q_bDone := FALSE;
q_bError := FALSE;
_bStartInput := FALSE; _bStartHolding := FALSE; _bStartWrite := FALSE; _bStartMulti := FALSE;
_rtExecute(CLK := i_bExecute);
IF _rtExecute.Q AND NOT q_bBusy THEN
	q_nErrorId := 0;
	IF i_sIpAddr = '' OR i_nPort = 0 OR i_nQuantity = 0 OR i_nQuantity > 125 THEN
		q_bDone := TRUE; q_bError := TRUE; q_nErrorId := 16#F001;
	ELSIF (i_nFunction = 6 AND (NOT GVL_PARAM.UPS_CONTROL_ENABLED OR NOT i_bWritePermit OR i_nQuantity <> 1))
		OR (i_nFunction = 16 AND (NOT GVL_PARAM.UPS_CONTROL_ENABLED OR NOT i_bWritePermit OR i_nQuantity > 3)) THEN
		q_bDone := TRUE; q_bError := TRUE; q_nErrorId := 16#F002;
	ELSIF i_nFunction <> 3 AND i_nFunction <> 4 AND i_nFunction <> 6 AND i_nFunction <> 16 THEN
		q_bDone := TRUE; q_bError := TRUE; q_nErrorId := 16#F003;
	ELSE
		_sIpAddr:=i_sIpAddr; _nPort:=i_nPort; _nUnitId:=i_nUnitId;
		_tTimeout:=i_tTimeout; _nAddress:=i_nAddress; _wValue:=i_wValue; _awValues:=i_awValues;
		_nFunction := i_nFunction; _nQuantity := i_nQuantity; q_bBusy := TRUE;
		_bStartInput := _nFunction = 4; _bStartHolding := _nFunction = 3; _bStartWrite := _nFunction = 6;
		_bStartMulti := _nFunction = 16;
	END_IF
END_IF
// Call all instances every scan, also while disabled, to drain an in-flight transaction.
_fbInput(sIPAddr:=_sIpAddr,nTCPPort:=_nPort,nUnitID:=_nUnitId,nMBAddr:=_nAddress,nQuantity:=_nQuantity,
	cbLength:=SIZEOF(q_awData),pDestAddr:=ADR(q_awData),tTimeout:=_tTimeout,bExecute:=_bStartInput);
_fbHolding(sIPAddr:=_sIpAddr,nTCPPort:=_nPort,nUnitID:=_nUnitId,nMBAddr:=_nAddress,nQuantity:=_nQuantity,
	cbLength:=SIZEOF(q_awData),pDestAddr:=ADR(q_awData),tTimeout:=_tTimeout,bExecute:=_bStartHolding);
_fbSingle(sIPAddr:=_sIpAddr,nTCPPort:=_nPort,nUnitID:=_nUnitId,nMBAddr:=_nAddress,nValue:=_wValue,tTimeout:=_tTimeout,bExecute:=_bStartWrite);
_fbMulti(sIPAddr:=_sIpAddr,nTCPPort:=_nPort,nUnitID:=_nUnitId,nQuantity:=_nQuantity,nMBAddr:=_nAddress,
	cbLength:=WORD_TO_UDINT(_nQuantity)*2,pSrcAddr:=ADR(_awValues),tTimeout:=_tTimeout,bExecute:=_bStartMulti);
IF q_bBusy THEN
	CASE _nFunction OF
		4: IF NOT _fbInput.bBusy AND NOT _bStartInput THEN
				q_bDone := TRUE; q_bError := _fbInput.bError OR (_fbInput.cbRead <> WORD_TO_UDINT(_nQuantity)*2);
				q_nErrorId := _fbInput.nErrId; q_bBusy := FALSE; END_IF
		3: IF NOT _fbHolding.bBusy AND NOT _bStartHolding THEN
				q_bDone := TRUE; q_bError := _fbHolding.bError OR (_fbHolding.cbRead <> WORD_TO_UDINT(_nQuantity)*2);
				q_nErrorId := _fbHolding.nErrId; q_bBusy := FALSE; END_IF
		6: IF NOT _fbSingle.bBusy AND NOT _bStartWrite THEN
				q_bDone := TRUE; q_bError := _fbSingle.bError; q_nErrorId := _fbSingle.nErrId; q_bBusy := FALSE; END_IF
		16: IF NOT _fbMulti.bBusy AND NOT _bStartMulti THEN
				q_bDone := TRUE; q_bError := _fbMulti.bError; q_nErrorId := _fbMulti.nErrId; q_bBusy := FALSE; END_IF
	END_CASE
	IF q_bDone AND q_bError AND q_nErrorId = 0 THEN q_nErrorId := 16#F004; END_IF
END_IF

END_FUNCTION_BLOCK

// ---- 20_Module/Ups/F_UpsNextSeq.TcPOU
FUNCTION F_UpsNextSeq : UDINT
VAR_INPUT i_nSeq : UDINT; END_VAR

IF i_nSeq = 16#FFFFFFFF THEN F_UpsNextSeq := 1;
ELSE F_UpsNextSeq := i_nSeq + 1; END_IF

END_FUNCTION

// ---- 20_Module/Virtual/FB_MeterSim.TcPOU
FUNCTION_BLOCK FB_MeterSim EXTENDS FB_DeviceBase IMPLEMENTS I_Meter		// 가상 계측기 (시험용)
VAR_INPUT
	i_fP			: REAL;					// kW (방전 +). PRG_SimLink가 넣음
	i_fQ			: REAL;					// kvar
	i_fVPhase		: REAL := 13221.0;		// V, 상전압
	i_fHz			: REAL := 60.0;
	i_bForceInvalid	: BOOL;			// 시험: 접속점 P/Q 계측 무효 (값·통신·전압·주파수는 유지)
END_VAR
VAR
	_stMeter		: ST_MeterState;
END_VAR

PROPERTY MeterState : ST_MeterState
GET
MeterState := _stMeter;
END_GET
END_PROPERTY

METHOD M_Cycle
VAR
	k		: UINT;
END_VAR
IF M_IsReadTime() THEN		// 읽기 주기마다 응답한 것으로 봄
	M_MarkAlive();
END_IF
M_UpdateComm();

_stMeter.bComm			:= _bComm;
_stMeter.stP.fValue		:= i_fP;
_stMeter.stP.bValid		:= NOT i_bForceInvalid;
_stMeter.stQ.fValue		:= i_fQ;
_stMeter.stQ.bValid		:= NOT i_bForceInvalid;
_stMeter.stV.fValue		:= i_fVPhase;
_stMeter.stV.bValid		:= TRUE;
FOR k := 1 TO 3 DO
	_stMeter.astV[k].fValue	:= i_fVPhase;
	_stMeter.astV[k].bValid	:= TRUE;
END_FOR
_stMeter.stF.fValue		:= i_fHz;
_stMeter.stF.bValid		:= TRUE;
END_METHOD

END_FUNCTION_BLOCK

// ---- 20_Module/Driver/Sebang/FB_SebangUps.TcPOU
FUNCTION_BLOCK FB_SebangUps EXTENDS FB_DeviceBase IMPLEMENTS I_Ups

VAR_INPUT
	i_bEnable : BOOL;
	i_sIpAddr : STRING(15);
	i_nPort : UINT := 502;
	i_nUnitId : BYTE := 1;
	i_tTimeout : TIME := T#1S;
	i_bWritePermit : BOOL; // site dispatcher: config OK AND active PLC
	i_bBlockStart : BOOL; // 2026-11-17: UPS 고장·e-stop 중 (MAIN이 보고 Status b2 OR b3로 줌). 시작 명령·설정 쓰기를 대기열에 넣지 않고, 이미 들어간 것도 뺌
END_VAR
VAR_OUTPUT
	q_eRequestResult : E_UpsResult;
	q_nTransportError : UDINT;
END_VAR
VAR
	_fbJob : FB_UpsModbusJob;
	_bLaunch : BOOL;
	_bCurrentWrite : BOOL;
	_bDiscardResponse : BOOL; // response started before a disable must not complete a new snapshot
	_nFunction : UINT;
	_nAddress : WORD;
	_nQuantity : WORD;
	_wValue : WORD;
	_bPendingWrite : BOOL;
	_nPendingAddress : WORD;
	_wPendingValue : WORD;
	_nPoll : UINT;
	_nCopy : UINT;
	_bReadDue : BOOL;
	_bCycle : BOOL; // 2026-11-23 한 바퀴(요청 4개) 읽는 중. i_tReadPeriod마다 시작해 4개를 연달아 읽음 (명세 DV-04 v2.46)
END_VAR

VAR_OUTPUT
	q_stRaw : ST_UpsRaw;
	q_stState : ST_UpsState;
END_VAR
VAR
	_stWork : ST_UpsRaw;
	_nSampleSeq : UDINT;
END_VAR

METHOD M_Cycle
_bReadDue := M_IsReadTime();
IF _bReadDue THEN _bCycle:=TRUE; END_IF // 한 바퀴 시작 (명세 DV-04 v2.46: 주기 = 한 바퀴)
IF NOT i_bEnable THEN
	_bDiscardResponse:=_bDiscardResponse OR _fbJob.q_bBusy;
	_bLaunch:=FALSE;
END_IF
IF NOT i_bEnable OR NOT i_bWritePermit OR NOT GVL_PARAM.UPS_CONTROL_ENABLED THEN
	_bPendingWrite := FALSE;
	// A queued but not yet started FC06 must not survive a gate transition.
	IF _bLaunch AND _bCurrentWrite THEN _bLaunch := FALSE; END_IF
END_IF
// 2026-11-17: 대기 중에 고장·e-stop이 생기면 시작 명령(켜기·시작)과 설정 쓰기를 뺀다. 끄기·취소·리셋(101,103,105,107,109,113,117,119,121,123,125,100)은 그대로
IF i_bBlockStart THEN
	IF _bPendingWrite THEN
		CASE _nPendingAddress OF
			7..64, 102, 104, 106, 108, 110, 111, 112, 114, 115, 116, 118, 120, 122, 124:
				_bPendingWrite := FALSE;
				q_eRequestResult := E_UpsResult.BadRequest;
		END_CASE
	END_IF
	IF _bLaunch AND _bCurrentWrite THEN
		CASE _nAddress OF
			7..64, 102, 104, 106, 108, 110, 111, 112, 114, 115, 116, 118, 120, 122, 124:
				_bLaunch := FALSE;
				_bCurrentWrite := FALSE;
				q_eRequestResult := E_UpsResult.BadRequest;
		END_CASE
	END_IF
END_IF
_fbJob(i_sIpAddr:=i_sIpAddr,i_nPort:=i_nPort,i_nUnitId:=i_nUnitId,i_tTimeout:=i_tTimeout,
	i_bExecute:=_bLaunch,i_bWritePermit:=i_bWritePermit AND i_bEnable,
	i_nFunction:=_nFunction,i_nAddress:=_nAddress,i_nQuantity:=_nQuantity,i_wValue:=_wValue);
_bLaunch := FALSE;
IF _fbJob.q_bDone THEN
	q_nTransportError := _fbJob.q_nErrorId;
	IF _bCurrentWrite THEN M_MarkWriteResult(NOT _fbJob.q_bError); END_IF
END_IF

IF _fbJob.q_bDone AND _bDiscardResponse THEN
	_bDiscardResponse:=FALSE; _nPoll:=0; _bCycle:=FALSE;
ELSIF _fbJob.q_bDone AND NOT _bCurrentWrite THEN
	IF _fbJob.q_bError THEN _nPoll:=0; _bCycle:=FALSE; // 다음 주기에 처음부터
	ELSE
		CASE _nPoll OF
			0: FOR _nCopy:=0 TO 34 DO _stWork.awInput[_nCopy]:=_fbJob.q_awData[_nCopy]; END_FOR
			1: FOR _nCopy:=0 TO 15 DO _stWork.awInput[_nCopy+38]:=_fbJob.q_awData[_nCopy]; END_FOR
			2: FOR _nCopy:=0 TO 11 DO _stWork.awParam[_nCopy]:=_fbJob.q_awData[_nCopy]; END_FOR
			3: FOR _nCopy:=0 TO 16 DO _stWork.awParam[_nCopy+50]:=_fbJob.q_awData[_nCopy]; END_FOR
		END_CASE
		IF _nPoll=3 THEN
			q_stRaw:=_stWork; _nSampleSeq:=F_UpsNextSeq(_nSampleSeq); M_MarkAlive(); _nPoll:=0; _bCycle:=FALSE;
		ELSE _nPoll:=_nPoll+1; END_IF
	END_IF
END_IF
M_UpdateComm();
q_stState:=F_DecodeSebangUps(q_stRaw);
q_stState.bComm:=_bComm AND i_bEnable;
q_stState.bValid:=q_stState.bComm AND _nSampleSeq<>0;
q_stState.nSampleSeq:=_nSampleSeq;
q_stState.bWriteFail:=_bWriteFail;
IF NOT _fbJob.q_bBusy AND NOT _fbJob.q_bDone AND i_bEnable AND i_sIpAddr<>'' THEN
IF _bPendingWrite THEN
	_nFunction:=6; _nAddress:=_nPendingAddress; _nQuantity:=1; _wValue:=_wPendingValue;
	_bCurrentWrite:=TRUE; _bPendingWrite:=FALSE; _bLaunch:=TRUE;
ELSIF _bCycle THEN // 한 바퀴 안에서는 앞 요청이 끝나면 바로 다음 요청 (쓰기가 있으면 쓰기 먼저)
	_bCurrentWrite:=FALSE;

	CASE _nPoll OF
		0: _nFunction:=4; _nAddress:=0; _nQuantity:=35;
		1: _nFunction:=4; _nAddress:=38; _nQuantity:=16;
		2: _nFunction:=3; _nAddress:=0; _nQuantity:=12;
		3: _nFunction:=3; _nAddress:=50; _nQuantity:=17;
	END_CASE
	_bLaunch:=TRUE;
	END_IF
END_IF
IF NOT i_bEnable THEN _nSampleSeq:=0; _nPoll:=0; _bLaunch:=FALSE; _bCycle:=FALSE; END_IF
END_METHOD

PROPERTY UpsState : ST_UpsState
GET
UpsState:=q_stState;
END_GET
END_PROPERTY

METHOD PRIVATE M_QueueWrite : BOOL
VAR_INPUT i_nAddress : WORD; i_wValue : WORD; END_VAR
q_eRequestResult := E_UpsResult.Disabled;
IF NOT GVL_PARAM.UPS_CONTROL_ENABLED OR NOT i_bWritePermit OR NOT i_bEnable THEN RETURN; END_IF
IF i_bBlockStart THEN // 2026-11-17: 고장·e-stop 중 시작 명령·설정 쓰기는 받지 않음
	CASE i_nAddress OF
		7..64, 102, 104, 106, 108, 110, 111, 112, 114, 115, 116, 118, 120, 122, 124:
			q_eRequestResult := E_UpsResult.BadRequest;
			RETURN;
	END_CASE
END_IF
q_eRequestResult := E_UpsResult.CommUnavailable;
IF NOT _bComm THEN RETURN; END_IF
q_eRequestResult := E_UpsResult.Busy;
IF _bPendingWrite OR _bCurrentWrite AND (_fbJob.q_bBusy OR _bLaunch) THEN RETURN; END_IF
_nPendingAddress := i_nAddress; _wPendingValue := i_wValue; _bPendingWrite := TRUE;
q_eRequestResult := E_UpsResult.Accepted;
M_QueueWrite := TRUE;
END_METHOD

METHOD M_RequestCommand : BOOL
VAR_INPUT i_eCommand : E_UpsCommand; END_VAR
CASE i_eCommand OF
	E_UpsCommand.Reset,
	E_UpsCommand.BuzzerStop,
	E_UpsCommand.RectifierOn,
	E_UpsCommand.RectifierOff,
	E_UpsCommand.InverterOn,
	E_UpsCommand.InverterOff,
	E_UpsCommand.BbcOn,
	E_UpsCommand.BbcOff,
	E_UpsCommand.ToInverter,
	E_UpsCommand.ToBypass,
	E_UpsCommand.FloatCharge,
	E_UpsCommand.EqualCharge,
	E_UpsCommand.AutoOn,
	E_UpsCommand.AutoOff,
	E_UpsCommand.EmergencyDischarge,
	E_UpsCommand.PeriodicDischarge,
	E_UpsCommand.PulseDischarge,
	E_UpsCommand.CancelDischarge,
	E_UpsCommand.TrickleOn,
	E_UpsCommand.TrickleOff,
	E_UpsCommand.TemperatureOn,
	E_UpsCommand.TemperatureOff,
	E_UpsCommand.EcoOn,
	E_UpsCommand.EcoOff,
	E_UpsCommand.PrltOn,
	E_UpsCommand.PrltOff:
	M_RequestCommand:=M_QueueWrite(INT_TO_WORD(TO_INT(i_eCommand)),16#0055);
ELSE q_eRequestResult:=E_UpsResult.Unsupported;
END_CASE
END_METHOD

METHOD M_SetParameter : BOOL
// Explicit RAW register value only. 57~59 allowed since 2026-11-16 (spec v2.14: H58/H59 = voltage or SOC by H57). 62 still rejected (scale O-11).
VAR_INPUT i_nAddress : WORD; i_wRawValue : WORD; END_VAR
CASE i_nAddress OF
	7,8,10,50,51,52,53,54,55,56,57,58,59,60,61,63,64:
		M_SetParameter:=M_QueueWrite(i_nAddress,i_wRawValue);
ELSE q_eRequestResult:=E_UpsResult.Unsupported;
END_CASE
END_METHOD

METHOD M_CheckSet : WSTRING(63)
M_CheckSet:="";
IF i_bEnable THEN
	IF i_sIpAddr='' OR i_nPort=0 THEN M_CheckSet:="TCP endpoint missing";
	ELSIF i_tReadPeriod<=T#0MS OR i_tTimeout<=T#0MS OR i_tCommTimeout<=i_tReadPeriod THEN M_CheckSet:="Invalid timing";
	END_IF
END_IF
END_METHOD

END_FUNCTION_BLOCK

// ---- 20_Module/Driver/Sebang/F_DecodeSebangUps.TcPOU
FUNCTION F_DecodeSebangUps : ST_UpsState
VAR_INPUT i_stRaw : ST_UpsRaw; END_VAR
VAR n : UINT; END_VAR

// UPS Metering Data 주소 순서
F_DecodeSebangUps.fInputVoltageRV := WORD_TO_REAL(i_stRaw.awInput[0])*0.1; // 0. 입력 선간 전압 R (V)
F_DecodeSebangUps.fInputVoltageSV := WORD_TO_REAL(i_stRaw.awInput[1])*0.1; // 1. 입력 선간 전압 S (V)
F_DecodeSebangUps.fInputVoltageTV := WORD_TO_REAL(i_stRaw.awInput[2])*0.1; // 2. 입력 선간 전압 T (V)
F_DecodeSebangUps.fInputFrequencyHz := WORD_TO_REAL(i_stRaw.awInput[3])*0.1; // 3. 입력 주파수 (Hz)
F_DecodeSebangUps.fInputCurrentRA := WORD_TO_REAL(i_stRaw.awInput[4])*0.1; // 4. 입력 전류 R (A)
F_DecodeSebangUps.fInputCurrentSA := WORD_TO_REAL(i_stRaw.awInput[5])*0.1; // 5. 입력 전류 S (A)
F_DecodeSebangUps.fInputCurrentTA := WORD_TO_REAL(i_stRaw.awInput[6])*0.1; // 6. 입력 전류 T (A)
F_DecodeSebangUps.fInverterVoltageRV := WORD_TO_REAL(i_stRaw.awInput[7])*0.1; // 7. 인버터 선간 전압 R (V)
F_DecodeSebangUps.fInverterVoltageSV := WORD_TO_REAL(i_stRaw.awInput[8])*0.1; // 8. 인버터 선간 전압 S (V)
F_DecodeSebangUps.fInverterVoltageTV := WORD_TO_REAL(i_stRaw.awInput[9])*0.1; // 9. 인버터 선간 전압 T (V)
F_DecodeSebangUps.fInverterCurrentRA := WORD_TO_REAL(i_stRaw.awInput[10])*0.1; // 10. 인버터 전류 R (A)
F_DecodeSebangUps.fInverterCurrentSA := WORD_TO_REAL(i_stRaw.awInput[11])*0.1; // 11. 인버터 전류 S (A)
F_DecodeSebangUps.fInverterCurrentTA := WORD_TO_REAL(i_stRaw.awInput[12])*0.1; // 12. 인버터 전류 T (A)
F_DecodeSebangUps.fBypassVoltageRV := WORD_TO_REAL(i_stRaw.awInput[13])*0.1; // 13. 바이패스 선간 전압 R (V)
F_DecodeSebangUps.fBypassVoltageSV := WORD_TO_REAL(i_stRaw.awInput[14])*0.1; // 14. 바이패스 선간 전압 S (V)
F_DecodeSebangUps.fBypassVoltageTV := WORD_TO_REAL(i_stRaw.awInput[15])*0.1; // 15. 바이패스 선간 전압 T (V)
F_DecodeSebangUps.fBypassFrequencyHz := WORD_TO_REAL(i_stRaw.awInput[16])*0.1; // 16. 바이패스 주파수 (Hz)
F_DecodeSebangUps.fOutputVoltageRV := WORD_TO_REAL(i_stRaw.awInput[17])*0.1; // 17. 출력 선간 전압 R (V)
F_DecodeSebangUps.fOutputVoltageSV := WORD_TO_REAL(i_stRaw.awInput[18])*0.1; // 18. 출력 선간 전압 S (V)
F_DecodeSebangUps.fOutputVoltageTV := WORD_TO_REAL(i_stRaw.awInput[19])*0.1; // 19. 출력 선간 전압 T (V)
F_DecodeSebangUps.fOutputFrequencyHz := WORD_TO_REAL(i_stRaw.awInput[20])*0.1; // 20. 출력 주파수 (Hz)
F_DecodeSebangUps.fOutputCurrentRA := WORD_TO_REAL(i_stRaw.awInput[21])*0.1; // 21. 출력 전류 R (A)
F_DecodeSebangUps.fOutputCurrentSA := WORD_TO_REAL(i_stRaw.awInput[22])*0.1; // 22. 출력 전류 S (A)
F_DecodeSebangUps.fOutputCurrentTA := WORD_TO_REAL(i_stRaw.awInput[23])*0.1; // 23. 출력 전류 T (A)
F_DecodeSebangUps.fDcLinkVoltageV := F_UpsSignedWord(i_stRaw.awInput[24])*0.1; // 24. DC 링크 전압 (V)
F_DecodeSebangUps.fDcLinkHighVoltageV := F_UpsSignedWord(i_stRaw.awInput[25])*0.1; // 25. DC 링크 상단 전압 (V)
F_DecodeSebangUps.fDcLinkLowVoltageV := F_UpsSignedWord(i_stRaw.awInput[26])*0.1; // 26. DC 링크 하단 전압 (V)
F_DecodeSebangUps.fBatteryVoltageV := F_UpsSignedWord(i_stRaw.awInput[27])*0.1; // 27. 배터리 전압 (V)
F_DecodeSebangUps.fBatteryCurrentA := F_UpsSignedWord(i_stRaw.awInput[28])*0.1; // 28. 배터리 전류 (A)
F_DecodeSebangUps.fMpiCurrentAA := F_UpsSignedWord(i_stRaw.awInput[29])*0.1; // 29. MPI A상 전류 (A)
F_DecodeSebangUps.fMpiCurrentBA := F_UpsSignedWord(i_stRaw.awInput[30])*0.1; // 30. MPI B상 전류 (A)
F_DecodeSebangUps.fMpiCurrentCA := F_UpsSignedWord(i_stRaw.awInput[31])*0.1; // 31. MPI C상 전류 (A)
F_DecodeSebangUps.fInputApparentPowerKva := F_UpsSignedWord(i_stRaw.awInput[32])*0.1; // 32. 입력 피상 전력 (kVA)
F_DecodeSebangUps.fOutputApparentPowerKva := F_UpsSignedWord(i_stRaw.awInput[33])*0.1; // 33. 출력 피상 전력 (kVA)
F_DecodeSebangUps.fOutputActivePowerKw := F_UpsSignedWord(i_stRaw.awInput[34])*0.1; // 34. 출력 유효 전력 (kW)
F_DecodeSebangUps.fTemperature1C := F_UpsSignedWord(i_stRaw.awInput[38])*0.1; // 38. 온도 1 (℃)
F_DecodeSebangUps.fTemperature2C := F_UpsSignedWord(i_stRaw.awInput[39])*0.1; // 39. 온도 2 (℃)
F_DecodeSebangUps.fTemperature3C := F_UpsSignedWord(i_stRaw.awInput[40])*0.1; // 40. 온도 3 (℃)
F_DecodeSebangUps.fTemperature4C := F_UpsSignedWord(i_stRaw.awInput[41])*0.1; // 41. 온도 4 (℃)
F_DecodeSebangUps.fTemperature5C := F_UpsSignedWord(i_stRaw.awInput[42])*0.1; // 42. 온도 5 (℃)
F_DecodeSebangUps.fBatteryRoomTemperatureC := F_UpsSignedWord(i_stRaw.awInput[43])*0.1; // 43. 온도 6 / 배터리실 온도 (℃)
F_DecodeSebangUps.wInputAlarm := i_stRaw.awInput[44]; // 44. 입력 알람
F_DecodeSebangUps.wRectAlarm := i_stRaw.awInput[45]; // 45. 정류기 알람
F_DecodeSebangUps.wBbcAlarm := i_stRaw.awInput[46]; // 46. 배터리 컨버터 알람
F_DecodeSebangUps.wOutputAlarm := i_stRaw.awInput[47]; // 47. 출력 알람
F_DecodeSebangUps.wInverterAlarm := i_stRaw.awInput[48]; // 48. 인버터 알람
F_DecodeSebangUps.wBypassAlarm := i_stRaw.awInput[49]; // 49. 바이패스 알람
F_DecodeSebangUps.wStatus1 := i_stRaw.awInput[50]; // 50. 상태 워드 1
F_DecodeSebangUps.wStatus2 := i_stRaw.awInput[51]; // 51. 상태 워드 2
F_DecodeSebangUps.fHmiVersion := WORD_TO_REAL(i_stRaw.awInput[52])*0.1; // 52. HMI 버전
F_DecodeSebangUps.fDspVersion := WORD_TO_REAL(i_stRaw.awInput[53])*0.1; // 53. DSP 버전

F_DecodeSebangUps.nBatMode := WORD_TO_UINT(SHR(i_stRaw.awInput[50],8) AND 16#0007);
F_DecodeSebangUps.bRectOn := i_stRaw.awInput[45].11;
F_DecodeSebangUps.bRectNormal := i_stRaw.awInput[45].12;
F_DecodeSebangUps.bBbcOn := i_stRaw.awInput[46].12;
F_DecodeSebangUps.bBbcNormal := i_stRaw.awInput[46].13;
F_DecodeSebangUps.bInverterOn := i_stRaw.awInput[48].6;
F_DecodeSebangUps.bInverterNormal := i_stRaw.awInput[48].14;
F_DecodeSebangUps.bOnBypass := i_stRaw.awInput[48].12;
F_DecodeSebangUps.bOnInverter := i_stRaw.awInput[48].13;
F_DecodeSebangUps.bTemperatureEnabled := i_stRaw.awInput[51].2;
F_DecodeSebangUps.bBmsMinor := i_stRaw.awInput[51].10;
F_DecodeSebangUps.bBmsMajor := i_stRaw.awInput[51].11;
F_DecodeSebangUps.bEmergencyStop := i_stRaw.awInput[50].0;
FOR n:=0 TO 7 DO F_DecodeSebangUps.awAlarmStatus[n]:=i_stRaw.awInput[n+44]; END_FOR
F_DecodeSebangUps.wOpCode := i_stRaw.awParam[11]; // H11 OP-CODE (b3 Batt CB Trip, 명세 RD-UPS-01 v2.50)

END_FUNCTION

// ---- 20_Module/Common/FB_RuleBit.TcPOU
FUNCTION_BLOCK FB_RuleBit EXTENDS FB_ModuleBase IMPLEMENTS I_ProtectionRule, I_OutputRule		// 디지털 접점 하나 → 조건 (화재·연기·비상정지·문 열림 등). 보호 규칙·출력 규칙 어느 쪽으로도 등록
VAR_INPUT
	i_ipAux			: I_AuxDevice;		// 읽을 보조 장비 (선언 때 지정)
	i_nPoint		: UINT;				// 디지털 입력 점 번호
	i_stSet			: ST_RuleBitSet;	// 설정: b접점, 통신 끊김 시 조건 (MAIN이 GVL_PERSIST.g_stModuleSet 칸을 매 스캔 넘김. 안 넘기면 기본값)
END_VAR
VAR
	_bCond			: BOOL;
END_VAR

METHOD M_Evaluate : BOOL		// 보호 규칙으로 판단 (범위·대상과 관계없이 접점 하나)
VAR_INPUT
	i_stView	: ST_ProtView;
END_VAR
M_Evaluate := M_Check(i_fThreshold := i_stView.fThreshold);
END_METHOD

METHOD M_Check : BOOL		// 출력 규칙으로 판단. 보호 판단도 이것을 씀
VAR_INPUT
	i_fThreshold	: REAL;			// 안 씀
END_VAR
IF i_ipAux = 0 THEN
	_bCond := FALSE;
ELSIF NOT i_ipAux.Comm THEN
	_bCond := i_stSet.bOnCommLoss;
ELSE
	_bCond := i_ipAux.M_GetBit(i_nPoint) XOR i_stSet.bInvert;
END_IF
M_Check := _bCond;
END_METHOD

END_FUNCTION_BLOCK

// ---- 20_Module/Driver/Autonics/FB_AutonicsThd.TcPOU
FUNCTION_BLOCK FB_AutonicsThd EXTENDS FB_DeviceBase IMPLEMENTS I_AuxDevice		// 오토닉스 THD 온습도계 (Modbus RTU, 한 줄에 국번 1..n), 읽기 전용
(* ---------------------------------------------------------------
   기반: Helios FB_ThdAutonics_Chain (PRG_Sensor에서 쓰던 것). 동작만 옮기고 PmsStd 드라이버 형식으로 다시 씀. 2026-11-09
   통신: 시리얼 단자(EL6022 채널 하나, 사용자 2026-11-09 회사 표준)를 ModbusRtuMaster_KL6x22B로. 단자 연결(InData·OutData)은 XAE I/O 화면에서 사람이 함
   읽기: 읽기 주기마다 센서 하나씩 돌아가며 Input Register(FC4)
     @MAP IR 0 S16 0.01 ℃  온도
     @MAP IR 1 S16 0.01 %  습도
   점 (I_AuxDevice)
     AI 2n-1 = 센서 n 온도 (℃), AI 2n = 센서 n 습도 (%). 센서 n이 i_tCommTimeout 동안 응답 없으면 bValid FALSE
     DI n    = 센서 n 통신 이상 (TRUE = 이상. Helios SensorStatus 1과 같음)
   센서는 GVL_PARAM.AUX_AI_MAX / 2개까지. 쓰기(DO·AO) 없음
   맵 미확보: Helios 현장 기종 기준. 실제 기종이 정해지면 주소·배율 확인
   --------------------------------------------------------------- *)
VAR_INPUT
	i_bEnable		: BOOL;					// FALSE면 통신하지 않음 (장비 미설치)
	i_nSensorCount	: UINT := 1;			// 국번 1..n 연속 (1..SENSOR_MAX)
	i_tTimeout		: TIME := T#1S;			// 응답 기다림 (Helios 5 s)
END_VAR
VAR
	_fbRtu			: ModbusRtuMaster_KL6x22B;
	_awRaw			: ARRAY[0..1] OF WORD;
	_bReadDue		: BOOL;					// 읽을 때가 됨 (매 스캔 M_IsReadTime)
	_bReading		: BOOL;
	_nUnit			: UINT;					// 지금 읽는 국번
	_nCount			: UINT;					// 쓰는 센서 수 (범위로 자른 i_nSensorCount)
	_afTemp			: ARRAY[1..SENSOR_MAX] OF REAL;
	_afHum			: ARRAY[1..SENSOR_MAX] OF REAL;
	_abReadOk		: ARRAY[1..SENSOR_MAX] OF BOOL;	// 이번 스캔에 응답 받음
	_abEverOk		: ARRAY[1..SENSOR_MAX] OF BOOL;	// 한 번이라도 응답 받음
	_abSensorOk		: ARRAY[1..SENSOR_MAX] OF BOOL;	// 센서 통신 정상
	_atonLoss		: ARRAY[1..SENSOR_MAX] OF TON;
	_nIdx			: UINT;
END_VAR
VAR CONSTANT
	SENSOR_MAX		: UINT := GVL_PARAM.AUX_AI_MAX / 2;
END_VAR

METHOD M_Cycle
_nCount := LIMIT(1, i_nSensorCount, SENSOR_MAX);

_bReadDue := M_IsReadTime();
IF NOT _bReading THEN
	IF i_bEnable AND _bReadDue THEN
		IF _nUnit >= _nCount THEN _nUnit := 1; ELSE _nUnit := _nUnit + 1; END_IF
		_fbRtu.ReadInputRegs(UnitID := UINT_TO_BYTE(_nUnit), Quantity := 2, MBAddr := 0,
			cbLength := SIZEOF(_awRaw), pMemoryAddr := ADR(_awRaw), Timeout := i_tTimeout, Execute := TRUE);
		_bReading := TRUE;
	END_IF
ELSE
	_fbRtu.ReadInputRegs(Execute := FALSE);	// 시작한 읽기는 끝까지 부름 (Helios와 같음)
	IF NOT _fbRtu.BUSY THEN
		IF NOT _fbRtu.Error AND i_bEnable THEN
			_afTemp[_nUnit]		:= INT_TO_REAL(WORD_TO_INT(_awRaw[0])) * 0.01;	// @MAP IR 0 S16 0.01 ℃
			_afHum[_nUnit]		:= INT_TO_REAL(WORD_TO_INT(_awRaw[1])) * 0.01;	// @MAP IR 1 S16 0.01 %
			_abReadOk[_nUnit]	:= TRUE;
			_abEverOk[_nUnit]	:= TRUE;
			M_MarkAlive();
		END_IF
		_bReading := FALSE;
	END_IF
END_IF

FOR _nIdx := 1 TO SENSOR_MAX DO
	_atonLoss[_nIdx](IN := NOT _abReadOk[_nIdx], PT := i_tCommTimeout);
	_abSensorOk[_nIdx]	:= i_bEnable AND _nIdx <= _nCount AND _abEverOk[_nIdx] AND NOT _atonLoss[_nIdx].Q;
	_abReadOk[_nIdx]	:= FALSE;
END_FOR
M_UpdateComm();
END_METHOD

METHOD M_GetBit : BOOL		// DI n = 센서 n 통신 이상
VAR_INPUT
	i_nPoint	: UINT;
END_VAR
IF i_nPoint >= 1 AND i_nPoint <= _nCount THEN
	M_GetBit := NOT _abSensorOk[i_nPoint];
END_IF
END_METHOD

METHOD M_GetValue : ST_Val		// AI 2n-1 = 센서 n 온도 (℃), AI 2n = 센서 n 습도 (%)
VAR_INPUT
	i_nPoint	: UINT;
END_VAR
VAR
	nSensor		: UINT;
END_VAR
nSensor := (i_nPoint + 1) / 2;
IF i_nPoint >= 1 AND nSensor <= _nCount THEN
	M_GetValue.fValue := SEL(i_nPoint MOD 2 = 1, _afHum[nSensor], _afTemp[nSensor]);
	M_GetValue.bValid := _abSensorOk[nSensor];
END_IF
END_METHOD

METHOD M_SetBit		// 출력 없음
VAR_INPUT
	i_nPoint	: UINT;
	i_bValue	: BOOL;
END_VAR
;
END_METHOD

METHOD M_SetValue		// 출력 없음
VAR_INPUT
	i_nPoint	: UINT;
	i_fValue	: REAL;
END_VAR
;
END_METHOD

PROPERTY Comm : BOOL
GET
Comm := _bComm AND i_bEnable;
END_GET
END_PROPERTY

END_FUNCTION_BLOCK

// ---- 20_Module/Driver/LS/FB_LsImd1000.TcPOU
FUNCTION_BLOCK FB_LsImd1000 EXTENDS FB_DeviceBase IMPLEMENTS I_AuxDevice		// LS IMD1000 절연감시장치(IMD) (Modbus TCP, RS485 게이트웨이 경유), 읽기 전용
(* ---------------------------------------------------------------
   기반: MESSIS(TC2) FB_LsIMD1000. 주소는 LS 맵으로 고침. 2026-11-09
   맵: 인터페이스\(MM-20210721) IMD1000 Modbus-Setting_v1_0_0.pdf (장비는 RS485 RTU 전용 → 현장은 RS485-TCP 게이트웨이, 사용자 결정)
   읽기 (프로토콜 주소, 0 기준 = 맵 Addr 열)
     측정: Input Register(FC4) 199부터 36개 (MESSIS와 같은 범위)
       @MAP IR 206 U16  기기 DI 입력 상태
       @MAP IR 209 U16  자가진단 Error #2
       @MAP IR 210 U16  절연저항 alarm 상태
       @MAP IR 211 U16  기기 & 계통 연결 상태
       @MAP IR 215 U16  Self Test 진행 상태
       @MAP IR 224~225 F32(앞 = 상위)  절연저항 kΩ
       MESSIS는 223~224를 읽어 한 칸 어긋나 있었다(223 = 커패시턴스 상태). 상위 워드가 맞아 값은 거의 같게 보였음
     설정: Holding Register(FC3) 40부터 8개, 측정 SET_EVERY번에 한 번
       @MAP HR 40~41 U32(앞 = 상위)  Ins. Alarm Pick-up kΩ
       @MAP HR 46~47 U32  Pre Alarm#1 Pick-up kΩ
   점 (I_AuxDevice). DI 2는 Bender ISO685 드라이버와 같은 "보호용 경보"
     AI 1 절연저항, 2 Ins. Alarm 설정값, 3 Pre Alarm#1 설정값
     DI 1 경고 (Pre#1 OR Pre#2), 2 절연 경보 (Ins. Alarm), 3 시험 중, 4 사전경고 (Pre#3), 5 기기 고장 (자가진단·Device), 6 계통 연결 이상, 7 접지(PE) 연결 이상
   쓰기 없음 (릴레이·Self Test 제어는 하지 않음)
   --------------------------------------------------------------- *)
VAR_INPUT
	i_bEnable		: BOOL;					// FALSE면 통신하지 않음 (장비 미설치)
	i_sIpAddr		: STRING(15);			// 게이트웨이 주소
	i_nPort			: UINT := 502;
	i_nUnitId		: BYTE := 1;			// IMD1000 국번 (장비 초기값 1)
	i_tTimeout		: TIME := T#1S;
END_VAR
VAR_OUTPUT
	q_stState		: ST_LsImd1000State;	// 읽은 값 (보고 매핑 FB_RptLsImd1000이 씀)
END_VAR
VAR
	_fbIr			: FB_MBReadInputRegs;	// 측정 (FC4)
	_fbHr			: FB_MBReadRegs;		// 설정 (FC3)
	_awIr			: ARRAY[0..35] OF WORD;	// IR 199..234
	_awSet			: ARRAY[0..7] OF WORD;	// HR 40..47
	_bReadDue		: BOOL;					// 읽을 때가 됨 (매 스캔 M_IsReadTime)
	_bReading		: BOOL;
	_bSetBlock		: BOOL;					// 이번 읽기가 설정 영역
	_bBusy			: BOOL;
	_bError			: BOOL;
	_nReadCnt		: UINT;					// 0이면 설정 영역을 읽음 (부팅 직후 먼저)
	_bMeasOk		: BOOL;					// 측정 영역을 한 번 이상 읽음
END_VAR
VAR CONSTANT
	IR_ADDR			: UINT := 199;
	IR_QTY			: UINT := 36;
	SET_ADDR		: UINT := 40;
	SET_QTY			: UINT := 8;
	SET_EVERY		: UINT := 10;			// 설정 영역은 읽기 10번에 한 번
END_VAR

ACTION A_MapMeas:
q_stState.wDiState		:= _awIr[7];		// @MAP IR 206
q_stState.wSelfDiag		:= _awIr[10];		// @MAP IR 209
q_stState.wAlarm		:= _awIr[11];		// @MAP IR 210
q_stState.wConnect		:= _awIr[12];		// @MAP IR 211
q_stState.wSelfTest		:= _awIr[16];		// @MAP IR 215
q_stState.fInsulation	:= F_WordsToReal(i_wHigh := _awIr[25], i_wLow := _awIr[26]);	// @MAP IR 224(상위)·225(하위) F32 kΩ
_bMeasOk := TRUE;
END_ACTION

ACTION A_MapSet:
q_stState.nInsPickup	:= SHL(WORD_TO_UDINT(_awSet[0]), 16) OR WORD_TO_UDINT(_awSet[1]);	// @MAP HR 40~41 U32
q_stState.nPre1Pickup	:= SHL(WORD_TO_UDINT(_awSet[6]), 16) OR WORD_TO_UDINT(_awSet[7]);	// @MAP HR 46~47 U32
q_stState.bSetValid		:= TRUE;
END_ACTION

METHOD M_Cycle
_bReadDue := M_IsReadTime();
IF NOT _bReading THEN
	IF i_bEnable AND i_sIpAddr <> '' AND _bReadDue THEN
		_bSetBlock := _nReadCnt = 0;
		IF _bSetBlock THEN
			_fbHr(sIPAddr := i_sIpAddr, nTCPPort := i_nPort, nUnitID := i_nUnitId,
				nQuantity := SET_QTY, nMBAddr := SET_ADDR, cbLength := SIZEOF(_awSet),
				pDestAddr := ADR(_awSet), tTimeout := i_tTimeout, bExecute := TRUE);
		ELSE
			_fbIr(sIPAddr := i_sIpAddr, nTCPPort := i_nPort, nUnitID := i_nUnitId,
				nQuantity := IR_QTY, nMBAddr := IR_ADDR, cbLength := SIZEOF(_awIr),
				pDestAddr := ADR(_awIr), tTimeout := i_tTimeout, bExecute := TRUE);
		END_IF
		_bReading := TRUE;
	END_IF
ELSE
	IF _bSetBlock THEN
		_fbHr(bExecute := FALSE);
		_bBusy := _fbHr.bBusy;
		_bError := _fbHr.bError;
	ELSE
		_fbIr(bExecute := FALSE);
		_bBusy := _fbIr.bBusy;
		_bError := _fbIr.bError;
	END_IF
	IF NOT _bBusy THEN
		IF NOT _bError AND i_bEnable THEN
			IF _bSetBlock THEN
				A_MapSet();
			ELSE
				A_MapMeas();
			END_IF
			M_MarkAlive();
		END_IF
		_nReadCnt := (_nReadCnt + 1) MOD SET_EVERY;
		_bReading := FALSE;
	END_IF
END_IF
M_UpdateComm();
q_stState.bValid := Comm AND _bMeasOk;
END_METHOD

METHOD M_GetBit : BOOL		// DI 1..7 (머리 주석). 통신 이상이면 FALSE (규칙 FB_RuleBit은 Comm으로 따로 판단)
VAR_INPUT
	i_nPoint	: UINT;
END_VAR
IF q_stState.bValid THEN
	CASE i_nPoint OF
		1: M_GetBit := q_stState.wAlarm.1 OR q_stState.wAlarm.2;
		2: M_GetBit := q_stState.wAlarm.0;
		3: M_GetBit := q_stState.wSelfTest = 1 OR q_stState.wDiState.0 OR q_stState.wDiState.1;
		4: M_GetBit := q_stState.wAlarm.3;
		5: M_GetBit := (q_stState.wSelfDiag AND 16#0007) <> 0 OR q_stState.wConnect.1;
		6: M_GetBit := q_stState.wConnect.2;
		7: M_GetBit := q_stState.wConnect.0;
	END_CASE
END_IF
END_METHOD

METHOD M_GetValue : ST_Val		// AI 1 절연저항 kΩ, 2 Ins. Alarm 설정값 kΩ, 3 Pre Alarm#1 설정값 kΩ
VAR_INPUT
	i_nPoint	: UINT;
END_VAR
CASE i_nPoint OF
	1:
		M_GetValue.fValue := q_stState.fInsulation;
		M_GetValue.bValid := q_stState.bValid;
	2:
		M_GetValue.fValue := UDINT_TO_REAL(q_stState.nInsPickup);
		M_GetValue.bValid := q_stState.bValid AND q_stState.bSetValid;
	3:
		M_GetValue.fValue := UDINT_TO_REAL(q_stState.nPre1Pickup);
		M_GetValue.bValid := q_stState.bValid AND q_stState.bSetValid;
END_CASE
END_METHOD

METHOD M_SetBit		// 출력 없음
VAR_INPUT
	i_nPoint	: UINT;
	i_bValue	: BOOL;
END_VAR
;
END_METHOD

METHOD M_SetValue		// 출력 없음
VAR_INPUT
	i_nPoint	: UINT;
	i_fValue	: REAL;
END_VAR
;
END_METHOD

PROPERTY Comm : BOOL
GET
Comm := _bComm AND i_bEnable;
END_GET
END_PROPERTY

END_FUNCTION_BLOCK

// ---- 20_Module/Common/F_WordsToReal.TcPOU
FUNCTION F_WordsToReal : REAL		// 레지스터 2개(IEEE754 float)를 REAL로. 앞 레지스터 = 상위 워드. 숫자가 아니면(NaN·무한) 0
(* 기반: Helios FNC_OLD_IEEE754·FNC_TO_IEEE754 (Bender ISO685, ACURA3700에서 앞 레지스터가 상위 워드). 2026-11-09 *)
VAR_INPUT
	i_wHigh		: WORD;		// 앞 레지스터 (상위 16비트)
	i_wLow		: WORD;		// 뒤 레지스터 (하위 16비트)
END_VAR
VAR
	dwRaw		: DWORD;
	fValue		: REAL;
END_VAR

dwRaw := SHL(WORD_TO_DWORD(i_wHigh), 16) OR WORD_TO_DWORD(i_wLow);
IF (dwRaw AND 16#7F800000) = 16#7F800000 THEN	// 지수부가 모두 1 = NaN·무한
	F_WordsToReal := 0.0;
ELSE
	MEMCPY(destAddr := ADR(fValue), srcAddr := ADR(dwRaw), n := 4);
	F_WordsToReal := fValue;
END_IF

END_FUNCTION

// ---- 20_Module/Driver/Rootech/FB_RootechAcuraIo.TcPOU
FUNCTION_BLOCK FB_RootechAcuraIo EXTENDS FB_DeviceBase IMPLEMENTS I_AuxDevice		// 루텍 ACURA3700 원격 I/O (Modbus TCP): 접점 입력·아날로그 입력 읽기 전용
(* ---------------------------------------------------------------
   기반: Helios FB_ACURA3700. Helios는 이 장치의 DI로 화재(열)·연기·가스 감지기 접점을 받았다. 동작만 옮기고 PmsStd 형식으로 다시 씀. 2026-11-09
   모듈 배치 (Helios와 같음, 물리 순서대로 모듈마다 레지스터 100개):
     DIO 모듈 = i_nStartAddr,  AI 모듈 = i_nStartAddr + 100.  Holding Register(FC3)
   읽기: 읽기 주기마다 DIO와 AI를 번갈아
     @MAP HR start+4..11   U16 -  DI ch1..8 상태 (0 = 꺼짐)
     @MAP HR start+16..17  U16 -  DO ch1..2 상태
     @MAP HR start+122..133 F32(앞 = 상위) -  AI ch1..6 변환값
   점 (I_AuxDevice)
     DI 1..8 = 접점 입력 ch1..8,  DI 9..10 = DO ch1..2 상태
     AI 1..6 = 아날로그 입력 ch1..6 변환값 (장치에 설정한 단위)
   쓰기(DO·AO) 없음
   맵 미확보: Helios 현장 기준. 실제 모듈 구성·주소는 현장에서 확인
   --------------------------------------------------------------- *)
VAR_INPUT
	i_bEnable		: BOOL;					// FALSE면 통신하지 않음 (장비 미설치)
	i_sIpAddr		: STRING(15);
	i_nPort			: UINT := 502;
	i_nUnitId		: BYTE := 1;
	i_nStartAddr	: UINT := 12100;		// 첫 모듈(DIO) 시작 주소
	i_tTimeout		: TIME := T#1S;
END_VAR
VAR
	_fbMbRead		: FB_MBReadRegs;
	_awDio			: ARRAY[0..41] OF WORD;
	_awAi			: ARRAY[0..45] OF WORD;
	_bReadDue		: BOOL;					// 읽을 때가 됨 (매 스캔 M_IsReadTime)
	_bReading		: BOOL;
	_bReadAi		: BOOL;					// 이번 읽기가 AI 모듈
	_abDi			: ARRAY[1..10] OF BOOL;
	_afAi			: ARRAY[1..6] OF REAL;
	_bDioOk			: BOOL;					// DIO 모듈을 한 번이라도 읽음
	_bAiOk			: BOOL;					// AI 모듈을 한 번이라도 읽음
	_nIdx			: UINT;
END_VAR

ACTION A_MapDio:
FOR _nIdx := 1 TO 8 DO
	_abDi[_nIdx] := _awDio[_nIdx + 3] <> 0;		// @MAP HR start+4..11 U16 DI ch1..8
END_FOR
_abDi[9]	:= _awDio[16] <> 0;					// @MAP HR start+16 U16 DO ch1 상태
_abDi[10]	:= _awDio[17] <> 0;					// @MAP HR start+17 U16 DO ch2 상태
END_ACTION

ACTION A_MapAi:
FOR _nIdx := 1 TO 6 DO
	_afAi[_nIdx] := F_WordsToReal(i_wHigh := _awAi[20 + 2 * _nIdx], i_wLow := _awAi[21 + 2 * _nIdx]);	// @MAP HR start+122+2(n-1) F32 AI chn
END_FOR
END_ACTION

METHOD M_Cycle
_bReadDue := M_IsReadTime();
IF NOT _bReading THEN
	IF i_bEnable AND i_sIpAddr <> '' AND _bReadDue THEN
		_bReadAi := NOT _bReadAi;
		IF _bReadAi THEN
			_fbMbRead(sIPAddr := i_sIpAddr, nTCPPort := i_nPort, nUnitID := i_nUnitId,
				nQuantity := 46, nMBAddr := i_nStartAddr + 100, cbLength := SIZEOF(_awAi),
				pDestAddr := ADR(_awAi), tTimeout := i_tTimeout, bExecute := TRUE);
		ELSE
			_fbMbRead(sIPAddr := i_sIpAddr, nTCPPort := i_nPort, nUnitID := i_nUnitId,
				nQuantity := 42, nMBAddr := i_nStartAddr, cbLength := SIZEOF(_awDio),
				pDestAddr := ADR(_awDio), tTimeout := i_tTimeout, bExecute := TRUE);
		END_IF
		_bReading := TRUE;
	END_IF
ELSE
	_fbMbRead(bExecute := FALSE);
	IF NOT _fbMbRead.bBusy THEN
		IF NOT _fbMbRead.bError AND i_bEnable THEN
			IF _bReadAi THEN
				A_MapAi();
				_bAiOk := TRUE;
			ELSE
				A_MapDio();
				_bDioOk := TRUE;
			END_IF
			M_MarkAlive();
		END_IF
		_bReading := FALSE;
	END_IF
END_IF
M_UpdateComm();
END_METHOD

METHOD M_GetBit : BOOL		// DI 1..8 = 접점 입력, 9..10 = DO 상태. 통신 이상이면 FALSE (규칙 FB_RuleBit은 Comm으로 따로 판단)
VAR_INPUT
	i_nPoint	: UINT;
END_VAR
IF i_nPoint >= 1 AND i_nPoint <= 10 AND Comm AND _bDioOk THEN
	M_GetBit := _abDi[i_nPoint];
END_IF
END_METHOD

METHOD M_GetValue : ST_Val		// AI 1..6 = 아날로그 입력 변환값
VAR_INPUT
	i_nPoint	: UINT;
END_VAR
IF i_nPoint >= 1 AND i_nPoint <= 6 THEN
	M_GetValue.fValue := _afAi[i_nPoint];
	M_GetValue.bValid := Comm AND _bAiOk;
END_IF
END_METHOD

METHOD M_SetBit		// 출력 없음 (DO는 읽기만)
VAR_INPUT
	i_nPoint	: UINT;
	i_bValue	: BOOL;
END_VAR
;
END_METHOD

METHOD M_SetValue		// 출력 없음
VAR_INPUT
	i_nPoint	: UINT;
	i_fValue	: REAL;
END_VAR
;
END_METHOD

PROPERTY Comm : BOOL
GET
Comm := _bComm AND i_bEnable;
END_GET
END_PROPERTY

END_FUNCTION_BLOCK

// ---- 20_Module/Driver/ITGuard/FB_ItGuardIeSx.TcPOU
FUNCTION_BLOCK FB_ItGuardIeSx EXTENDS FB_DeviceBase IMPLEMENTS I_AuxDevice		// ITGuard(이노튜브) IE-SX 이더넷 온습도계 (Modbus TCP), 읽기 전용
(* ---------------------------------------------------------------
   기반: MESSIS TC3 FB_IE_SX (광주첨단공장). 동작만 옮기고 PmsStd 형식으로 다시 씀. 2026-11-09
   읽기: Input Register(FC4) 0부터 5개 (MESSIS와 같음, Unit ID 1)
     @MAP IR 0  U16  mode
     @MAP IR 1  S16  센서1 = 온도 × 0.01 ℃
     @MAP IR 2  S16  센서2 = 습도 × 0.01 %
     @MAP IR 3·4 S16  센서3·4 (프로브 없으면 32767)
   2026-11-09 PC에서 읽어 확인: [0, 2418, 3545, 32767, 32767] → 24.18 ℃, 35.45 %
   센서 값 32767 = 프로브 없음으로 보고 무효 처리 (센서3·4가 비었을 때 이 값)
   점 (I_AuxDevice): AI 1 온도, AI 2 습도, DI 1 값 이상(통신 정상인데 프로브 무효)
   통신 이상: 응답 없이 i_tCommTimeout(기본 10초, MESSIS는 30초)
   쓰기 없음
   --------------------------------------------------------------- *)
VAR_INPUT
	i_bEnable		: BOOL;					// FALSE면 통신하지 않음 (장비 미설치)
	i_sIpAddr		: STRING(15);
	i_nPort			: UINT := 502;
	i_nUnitId		: BYTE := 1;
	i_tTimeout		: TIME := T#1S;
END_VAR
VAR_OUTPUT
	q_stState		: ST_TempHumState;		// 읽은 값 (보고 매핑 FB_RptTempHum이 씀)
END_VAR
VAR
	_fbIr			: FB_MBReadInputRegs;
	_awIr			: ARRAY[0..4] OF WORD;	// IR 0..4
	_bReadDue		: BOOL;
	_bReading		: BOOL;
	_bDataOk		: BOOL;					// 한 번이라도 읽음
	_bProbeOk		: BOOL;					// 온도·습도 값이 32767이 아님
END_VAR
VAR CONSTANT
	READ_QTY		: UINT := 5;
	NO_PROBE		: WORD := 16#7FFF;		// 프로브 없음
END_VAR

ACTION A_Map:
_bProbeOk		:= _awIr[1] <> NO_PROBE AND _awIr[2] <> NO_PROBE;
q_stState.fTemp	:= INT_TO_REAL(WORD_TO_INT(_awIr[1])) * 0.01;	// @MAP IR 1 S16 ×0.01 ℃
q_stState.fHum	:= INT_TO_REAL(WORD_TO_INT(_awIr[2])) * 0.01;	// @MAP IR 2 S16 ×0.01 %
_bDataOk := TRUE;
END_ACTION

METHOD M_Cycle
_bReadDue := M_IsReadTime();
IF NOT _bReading THEN
	IF i_bEnable AND i_sIpAddr <> '' AND _bReadDue THEN
		_fbIr(sIPAddr := i_sIpAddr, nTCPPort := i_nPort, nUnitID := i_nUnitId,
			nQuantity := READ_QTY, nMBAddr := 0, cbLength := SIZEOF(_awIr),
			pDestAddr := ADR(_awIr), tTimeout := i_tTimeout, bExecute := TRUE);
		_bReading := TRUE;
	END_IF
ELSE
	_fbIr(bExecute := FALSE);
	IF NOT _fbIr.bBusy THEN
		IF NOT _fbIr.bError AND i_bEnable THEN
			A_Map();
			M_MarkAlive();
		END_IF
		_bReading := FALSE;
	END_IF
END_IF
M_UpdateComm();
q_stState.bValid := Comm AND _bDataOk AND _bProbeOk;
END_METHOD

METHOD M_GetBit : BOOL		// DI 1 값 이상 (통신은 정상인데 프로브 값 무효)
VAR_INPUT
	i_nPoint	: UINT;
END_VAR
IF i_nPoint = 1 THEN
	M_GetBit := Comm AND _bDataOk AND NOT _bProbeOk;
END_IF
END_METHOD

METHOD M_GetValue : ST_Val		// AI 1 온도 ℃, AI 2 습도 %
VAR_INPUT
	i_nPoint	: UINT;
END_VAR
CASE i_nPoint OF
	1:
		M_GetValue.fValue := q_stState.fTemp;
		M_GetValue.bValid := q_stState.bValid;
	2:
		M_GetValue.fValue := q_stState.fHum;
		M_GetValue.bValid := q_stState.bValid;
END_CASE
END_METHOD

METHOD M_SetBit		// 출력 없음
VAR_INPUT
	i_nPoint	: UINT;
	i_bValue	: BOOL;
END_VAR
;
END_METHOD

METHOD M_SetValue		// 출력 없음
VAR_INPUT
	i_nPoint	: UINT;
	i_fValue	: REAL;
END_VAR
;
END_METHOD

PROPERTY Comm : BOOL
GET
Comm := _bComm AND i_bEnable;
END_GET
END_PROPERTY

END_FUNCTION_BLOCK

// ---- 20_Module/Driver/Woonyoung/FB_WoonyoungGfr.TcPOU
FUNCTION_BLOCK FB_WoonyoungGfr EXTENDS FB_DeviceBase IMPLEMENTS I_AuxDevice		// 운영(Woonyoung) WYGF-D08/12/16NC 디지털 지락검출계전기 (Modbus RTU), 읽기 전용
(* ---------------------------------------------------------------
   기반 없음(신규). 맵: 프로토콜 맵 v3\지락검출 계전기.pdf (사용설명서 PAC-00084 REV.5, 제5장). 2026-11-10
   용도: AC 회로 누전(지락) 감시. ZCT 영상변류기 방식이라 배터리 DC 전로 지락은 못 봄 (DC는 IMD)
   통신: EL6022 채널 하나를 ModbusRtuMaster_KL6x22B로 (사용자 2026-11-10). 단자 연결(InData·OutData)은 XAE I/O 화면에서 사람이 함
         장비: RS-485 8N1, 국번 1~32 (공장 출하 OFF → 장비 Serial Setup에서 켜야 응답), 9600/19200/38400 (출하 19200)
   읽기: 읽기 주기마다 Input Register(FC4) 0부터 2 + 회로 수
     @MAP IR 0      U16  시스템 상태 (b8 시험 모드, b4 LPF, b3 고감도 ZCT, b2 자동복귀, b1 부저, b0 50Hz)
     @MAP IR 1      U16  회로별 지락 (b0 = 1회로 … b15 = 16회로, 1 = Fault)
     @MAP IR 2~17   U16  회로 1~16 누설전류, × 0.01 A (예: 0x03E8 = 10 A)
   쓰지 않는 것: FC03 0~31 회로별 감도·동작시간 설정, FC03 32~51 사고 기록, FC05 0 사고 기록 지우기
   점 (I_AuxDevice)
     AI n = 회로 n 누설전류 (A)
     DI n = 회로 n 지락 (n = 1..회로 수), DI 17 = 시험 모드 (장비에서 Circuit Test 중)
   --------------------------------------------------------------- *)
VAR_INPUT
	i_bEnable		: BOOL;					// FALSE면 통신하지 않음 (장비 미설치)
	i_nUnitId		: UINT := 1;			// 장비 국번 (Serial Setup Port No.)
	i_nChannels		: UINT := 8;			// 회로 수: 8 (D08NC), 12 (D12NC), 16 (D16NC)
	i_tTimeout		: TIME := T#1S;			// 응답 기다림
END_VAR
VAR_OUTPUT
	q_wStatus		: WORD;					// IR 0 시스템 상태
	q_wFault		: WORD;					// IR 1 회로별 지락 비트
	q_afCurrent		: ARRAY[1..16] OF REAL;	// 회로별 누설전류 A
	q_bValid		: BOOL;					// 통신 정상이고 한 번 이상 읽음
END_VAR
VAR
	_fbRtu			: ModbusRtuMaster_KL6x22B;
	_awRaw			: ARRAY[0..17] OF WORD;	// IR 0..17
	_bReadDue		: BOOL;
	_bReading		: BOOL;
	_bDataOk		: BOOL;
	_nCh			: UINT;					// 쓰는 회로 수 (8·12·16 중 가까운 범위로 자름)
	_i				: UINT;
END_VAR
VAR CONSTANT
	CH_MAX			: UINT := 16;
	PT_TEST			: UINT := 17;			// DI 17 = 시험 모드
END_VAR

ACTION A_Map:
q_wStatus := _awRaw[0];				// @MAP IR 0
q_wFault := _awRaw[1];				// @MAP IR 1
FOR _i := 1 TO CH_MAX DO
	IF _i <= _nCh THEN
		q_afCurrent[_i] := WORD_TO_REAL(_awRaw[1 + _i]) * 0.01;	// @MAP IR 2~17 U16 ×0.01 A
	ELSE
		q_afCurrent[_i] := 0.0;
	END_IF
END_FOR
_bDataOk := TRUE;
END_ACTION

METHOD M_Cycle
_nCh := LIMIT(1, i_nChannels, CH_MAX);

_bReadDue := M_IsReadTime();
IF NOT _bReading THEN
	IF i_bEnable AND _bReadDue AND i_nUnitId >= 1 AND i_nUnitId <= 247 THEN
		_fbRtu.ReadInputRegs(UnitID := UINT_TO_BYTE(i_nUnitId), Quantity := 2 + _nCh, MBAddr := 0,
			cbLength := SIZEOF(_awRaw), pMemoryAddr := ADR(_awRaw), Timeout := i_tTimeout, Execute := TRUE);
		_bReading := TRUE;
	END_IF
ELSE
	_fbRtu.ReadInputRegs(Execute := FALSE);	// 시작한 읽기는 끝까지 부름
	IF NOT _fbRtu.BUSY THEN
		IF NOT _fbRtu.Error AND i_bEnable THEN
			A_Map();
			M_MarkAlive();
		END_IF
		_bReading := FALSE;
	END_IF
END_IF
M_UpdateComm();
q_bValid := Comm AND _bDataOk;
END_METHOD

METHOD M_GetBit : BOOL		// DI n = 회로 n 지락, DI 17 = 시험 모드. 통신 이상이면 FALSE (규칙 FB_RuleBit은 Comm으로 따로 판단)
VAR_INPUT
	i_nPoint	: UINT;
END_VAR
IF q_bValid THEN
	IF i_nPoint >= 1 AND i_nPoint <= _nCh THEN
		M_GetBit := (q_wFault AND SHL(WORD#1, i_nPoint - 1)) <> 0;
	ELSIF i_nPoint = PT_TEST THEN
		M_GetBit := q_wStatus.8;
	END_IF
END_IF
END_METHOD

METHOD M_GetValue : ST_Val		// AI n = 회로 n 누설전류 (A)
VAR_INPUT
	i_nPoint	: UINT;
END_VAR
IF i_nPoint >= 1 AND i_nPoint <= _nCh THEN
	M_GetValue.fValue := q_afCurrent[i_nPoint];
	M_GetValue.bValid := q_bValid;
END_IF
END_METHOD

METHOD M_SetBit		// 출력 없음
VAR_INPUT
	i_nPoint	: UINT;
	i_bValue	: BOOL;
END_VAR
;
END_METHOD

METHOD M_SetValue		// 출력 없음
VAR_INPUT
	i_nPoint	: UINT;
	i_fValue	: REAL;
END_VAR
;
END_METHOD

PROPERTY Comm : BOOL
GET
Comm := _bComm AND i_bEnable;
END_GET
END_PROPERTY

END_FUNCTION_BLOCK

// ---- 20_Module/Driver/Gasdna/FB_GasdnaAsd57.TcPOU
FUNCTION_BLOCK FB_GasdnaAsd57 EXTENDS FB_DeviceBase IMPLEMENTS I_AuxDevice		// 가스디엔에이 ASD-57 열연복합 감지기 (Modbus RTU), 읽기 전용
(* ---------------------------------------------------------------
   기반 없음(신규). 맵: 프로토콜 맵 v3\ASD-5x(모드 버스 프로토콜)_ver1.1(22_0922).pdf, 결선: ASD-57_매뉴얼.pdf. 2026-11-10
   통신: EL6022 채널 하나를 ModbusRtuMaster_KL6x22B로. 단자 연결(InData·OutData)은 XAE I/O 화면에서 사람이 함
         장비: RS-485 9600 bps 고정, 8N1, 국번 1~126 (출하 1). 흰 TX+, 파랑 TX-
         속도가 9600 고정이라 다른 속도 장비(지락계전기 출하 19200)와 한 채널에 묶지 않음
         응답 뒤 10 ms 이상 지나 다음 요청 (읽기 주기 1 s라 맞음)
   읽기: 읽기 주기마다 Holding Register(FC3) 0부터 9칸
     @MAP HR 0 (40001) U16  1 Color 연기 농도 0~1000, ×0.1 %
     @MAP HR 1 (40002) U16  2 Color 연기 농도 0~1000, ×0.01 (맵 표기 x.xx, 단위 표기 없음)
     @MAP HR 2 (40003) U16  온도 0~1000, ×0.1 ℃ (ASD-57 전용)
     @MAP HR 3 (40004) U16  알람 상태: 0 없음, 1 연기 (1·2 Color 모두 알람값 초과), 2 온도 (ASD-57 전용)
     @MAP HR 4 (40005) U16  1 Color 연기 알람값 (출하 80)
     @MAP HR 5 (40006) U16  2 Color 연기 알람값 (출하 170)
     @MAP HR 6 (40007) U16  온도 알람값 ×0.1 ℃ (출하 700 = 70.0 ℃)
     @MAP HR 7 (40008) U16  딜레이 ×10 ms (최대 1000 = 10 s)
     @MAP HR 8 (40009) U16  통신 국번
   쓰지 않는 것: FC6 HR 4~8 설정 바꾸기, HR 50 ZERO 교정(1234). 설정은 장비 출하값 그대로 (바꾸려면 사용자 결정)
   알람 상태 3(연기 + 온도)은 맵에 없음 → 비트로 봄 (b0 연기, b1 온도)
   점 (I_AuxDevice)
     AI 1 = 1 Color 연기 %, AI 2 = 2 Color 연기, AI 3 = 온도 ℃
     DI 1 = 연기 알람, DI 2 = 온도 알람
   --------------------------------------------------------------- *)
VAR_INPUT
	i_bEnable		: BOOL;					// FALSE면 통신하지 않음 (장비 미설치)
	i_nUnitId		: UINT := 1;			// 장비 국번 (HR 8)
	i_tTimeout		: TIME := T#1S;			// 응답 기다림
END_VAR
VAR_OUTPUT
	q_fSmoke1		: REAL;					// 1 Color 연기 농도 %
	q_fSmoke2		: REAL;					// 2 Color 연기 농도
	q_fTemp			: REAL;					// 온도 ℃
	q_wAlarm		: WORD;					// HR 3 알람 상태 원시값
	q_bSmokeAlarm	: BOOL;					// 연기 알람
	q_bTempAlarm	: BOOL;					// 온도 알람
	q_anSet			: ARRAY[4..8] OF UINT;	// HR 4~8 설정값 원시값 (알람값, 딜레이, 국번)
	q_bValid		: BOOL;					// 통신 정상이고 한 번 이상 읽음
END_VAR
VAR
	_fbRtu			: ModbusRtuMaster_KL6x22B;
	_awRaw			: ARRAY[0..8] OF WORD;	// HR 0..8
	_bReadDue		: BOOL;
	_bReading		: BOOL;
	_bDataOk		: BOOL;
	_i				: UINT;
END_VAR
VAR CONSTANT
	READ_QTY		: UINT := 9;
END_VAR

ACTION A_Map:
q_fSmoke1 := WORD_TO_REAL(_awRaw[0]) * 0.1;		// @MAP HR 0 ×0.1 %
q_fSmoke2 := WORD_TO_REAL(_awRaw[1]) * 0.01;	// @MAP HR 1 ×0.01
q_fTemp := WORD_TO_REAL(_awRaw[2]) * 0.1;		// @MAP HR 2 ×0.1 ℃
q_wAlarm := _awRaw[3];							// @MAP HR 3
q_bSmokeAlarm := q_wAlarm.0;
q_bTempAlarm := q_wAlarm.1;
FOR _i := 4 TO 8 DO
	q_anSet[_i] := WORD_TO_UINT(_awRaw[_i]);	// @MAP HR 4~8
END_FOR
_bDataOk := TRUE;
END_ACTION

METHOD M_Cycle
_bReadDue := M_IsReadTime();
IF NOT _bReading THEN
	IF i_bEnable AND _bReadDue AND i_nUnitId >= 1 AND i_nUnitId <= 126 THEN
		_fbRtu.ReadRegs(UnitID := UINT_TO_BYTE(i_nUnitId), Quantity := READ_QTY, MBAddr := 0,
			cbLength := SIZEOF(_awRaw), pMemoryAddr := ADR(_awRaw), Timeout := i_tTimeout, Execute := TRUE);
		_bReading := TRUE;
	END_IF
ELSE
	_fbRtu.ReadRegs(Execute := FALSE);	// 시작한 읽기는 끝까지 부름
	IF NOT _fbRtu.BUSY THEN
		IF NOT _fbRtu.Error AND i_bEnable THEN
			A_Map();
			M_MarkAlive();
		END_IF
		_bReading := FALSE;
	END_IF
END_IF
M_UpdateComm();
q_bValid := Comm AND _bDataOk;
END_METHOD

METHOD M_GetBit : BOOL		// DI 1 연기 알람, DI 2 온도 알람. 통신 이상이면 FALSE (규칙 FB_RuleBit은 Comm으로 따로 판단)
VAR_INPUT
	i_nPoint	: UINT;
END_VAR
IF q_bValid THEN
	CASE i_nPoint OF
		1: M_GetBit := q_bSmokeAlarm;
		2: M_GetBit := q_bTempAlarm;
	END_CASE
END_IF
END_METHOD

METHOD M_GetValue : ST_Val		// AI 1 연기1 %, AI 2 연기2, AI 3 온도 ℃
VAR_INPUT
	i_nPoint	: UINT;
END_VAR
CASE i_nPoint OF
	1: M_GetValue.fValue := q_fSmoke1;
	2: M_GetValue.fValue := q_fSmoke2;
	3: M_GetValue.fValue := q_fTemp;
ELSE
	RETURN;
END_CASE
M_GetValue.bValid := q_bValid;
END_METHOD

METHOD M_SetBit		// 출력 없음
VAR_INPUT
	i_nPoint	: UINT;
	i_bValue	: BOOL;
END_VAR
;
END_METHOD

METHOD M_SetValue		// 출력 없음
VAR_INPUT
	i_nPoint	: UINT;
	i_fValue	: REAL;
END_VAR
;
END_METHOD

PROPERTY Comm : BOOL
GET
Comm := _bComm AND i_bEnable;
END_GET
END_PROPERTY

END_FUNCTION_BLOCK

// ---- 20_Module/Virtual/FB_SrcTest.TcPOU
FUNCTION_BLOCK FB_SrcTest EXTENDS FB_SourceBase		// 시험 지령원: 온라인으로 값을 써서 시험
VAR_INPUT
	i_ePcsReq			: E_PcsCmd;		// PCS 요청. 쓰면 1스캔 요청으로 나가고 None으로 돌아감
	i_nPcsUnit			: UINT;			// 0 = 그룹 전체, n = 유닛 n
	i_eBatReq			: E_BatCmd;		// 배터리 요청 (Close / Open). 쓰면 1스캔 요청으로 나가고 None으로 돌아감
	i_nBatGroup			: UINT;			// 0 = 전체, n = 배터리 그룹 n
	i_bPSetActive		: BOOL;
	i_fPSet				: REAL;			// kW, 접속점 기준 (방전 +)
	i_bQSetActive		: BOOL;
	i_fQSet				: REAL;			// kvar, 접속점 기준 (공급 +)
	i_bPLimActive		: BOOL;			// 지령원 P 제한 시험
	i_fPMax				: REAL;			// kW
	i_fPMin				: REAL;
	i_bQLimActive		: BOOL;			// 지령원 Q 제한 시험
	i_fQMax				: REAL;			// kvar
	i_fQMin				: REAL;
	(* 유닛별 값 시험 (유닛 하나) *)
	i_nUnit				: UINT;			// 0 = 안 씀
	i_bUnitPSetActive	: BOOL;
	i_fUnitPSet			: REAL;			// kW, 유닛 출력
	i_bSend				: BOOL;			// 같은 값을 다시 보낼 때 TRUE (값을 바꾸면 자동으로 새 지령)
END_VAR

METHOD M_UpdateOutput : BOOL
VAR
	u		: UINT;
	stOld	: ST_SourceOutput;
END_VAR
stOld := _stOut;

_stOut.bPSetActive	:= i_bPSetActive;
_stOut.fPSet		:= i_fPSet;
_stOut.bQSetActive	:= i_bQSetActive;
_stOut.fQSet		:= i_fQSet;
_stOut.bPLimActive	:= i_bPLimActive;
_stOut.fPMax		:= i_fPMax;
_stOut.fPMin		:= i_fPMin;
_stOut.bQLimActive	:= i_bQLimActive;
_stOut.fQMax		:= i_fQMax;
_stOut.fQMin		:= i_fQMin;
IF i_ePcsReq <> E_PcsCmd.None THEN
	_stOut.stPcsReq.eCmd	:= i_ePcsReq;
	_stOut.stPcsReq.nUnit	:= i_nPcsUnit;
	i_ePcsReq				:= E_PcsCmd.None;
END_IF
IF i_eBatReq <> E_BatCmd.None THEN
	_stOut.stBatReq.eCmd		:= i_eBatReq;
	_stOut.stBatReq.nBatGroup	:= i_nBatGroup;
	i_eBatReq					:= E_BatCmd.None;
END_IF

FOR u := 1 TO GVL_PARAM.UNIT_COUNT DO
	_stOut.astUnit[u].bPSetActive := FALSE;
END_FOR
IF i_nUnit >= 1 AND i_nUnit <= GVL_PARAM.UNIT_COUNT THEN
	_stOut.astUnit[i_nUnit].bPSetActive	:= i_bUnitPSetActive;
	_stOut.astUnit[i_nUnit].fPSet		:= i_fUnitPSet;
END_IF
// 새 지령: 값이 바뀌었거나 i_bSend
// [결함 13 수정 2026-11-04: 값 비교를 비트로 (운전원이 NaN을 넣어도 여기서 멈추지 않고 고르기에서 이상값으로 거름). 원래 _stOut.fPSet <> stOld.fPSet, _stOut.fQSet <> stOld.fQSet, …fPSet <> stOld.astUnit[u].fPSet]
_stOut.bNewSet := i_bSend
	OR _stOut.bPSetActive <> stOld.bPSetActive OR F_RealChanged(_stOut.fPSet, stOld.fPSet)
	OR _stOut.bQSetActive <> stOld.bQSetActive OR F_RealChanged(_stOut.fQSet, stOld.fQSet);
FOR u := 1 TO GVL_PARAM.UNIT_COUNT DO
	_stOut.bNewSet := _stOut.bNewSet
		OR _stOut.astUnit[u].bPSetActive <> stOld.astUnit[u].bPSetActive
		OR F_RealChanged(_stOut.astUnit[u].fPSet, stOld.astUnit[u].fPSet);
END_FOR
i_bSend := FALSE;

M_UpdateOutput := TRUE;		// 시험용: 항상 살아 있음 (만료 없음)
END_METHOD

END_FUNCTION_BLOCK

// ---- 20_Module/ControlMode/FB_CmPeakCut.TcPOU
FUNCTION_BLOCK FB_CmPeakCut EXTENDS FB_CmTariffBase		// 제어 모드: 피크컷 (Messis PEAK_SHAVING_MODE). 15분 평균 수전이 목표를 넘지 않게 방전
// 우선순위: 자동 충전 시간 → 잔량 방전 시간 (잔량 방전과 피크 제어 중 큰 값, 방전 허용 시간에만) → 피크 제어 (방전 허용 시간에만). 휴일·시각 무효 → 0
// 방전은 모두 역송 방지 (공통 설정). 피크 제어량 계산은 FB_CmPeakCalc (통합 모드와 같음)
VAR_INPUT
	i_stSet		: ST_CmPeakCutSet;		// 설정 (A_PassModuleSet이 GVL_PERSIST.g_stModuleSet.stCmPeakCut을 매 스캔 넘김)
END_VAR
VAR_OUTPUT
	q_fPeakCtrl	: REAL;		// 진단: 피크 제어량 (kW, FB_CmPeakCalc)
	q_nRemainMin	: UINT;		// 진단: 15분 구간 남은 분
	q_fExceeded	: REAL;		// 진단: 구간 목표 초과 수전 누적 (kW·분)
	q_fLoad1m	: REAL;		// 진단: 직전 1분 평균 부하 (kW)
END_VAR
VAR
	_fbPeak		: FB_CmPeakCalc;
END_VAR

METHOD M_Enter
VAR_INPUT
	i_stView	: ST_CtrlModeView;
END_VAR
SUPER^.M_Enter(i_stView := i_stView);
_fbPeak.M_Reset();
END_METHOD

METHOD M_Calc : ST_CtrlModeOut
VAR_INPUT
	i_stView	: ST_CtrlModeView;
END_VAR
VAR
	nNow	: UINT;
	fP		: REAL;
	fRem	: REAL;
	nRsn	: UINT;
	bNoCap	: BOOL;
END_VAR
fP := 0.0;
_fbPeak(i_stSet := i_stSet.stPeak, i_fRevMargin := i_stCommon.stNoRev.fMargin, i_stView := i_stView);		// 휴일에도 평균은 셈
q_fPeakCtrl		:= _fbPeak.q_fCtrl;
q_nRemainMin	:= _fbPeak.q_nRemainMin;
q_fExceeded		:= _fbPeak.q_fExceeded;
q_fLoad1m		:= _fbPeak.q_fLoad1m;
IF M_Begin(i_stView := i_stView) THEN
	nNow := F_TimeHhmm(i_stTime := i_stView.stTime);
	IF i_stSet.stAutoChg.bUse AND F_InHhmmWindow(i_nNow := nNow, i_nStart := i_stSet.stAutoChg.nStart, i_nEnd := i_stSet.stAutoChg.nEnd) THEN
		// 1) 자동 충전 (Messis MT_auto_charge)
		fP			:= -M_AutoChg(i_stView := i_stView, i_stWin := i_stSet.stAutoChg, q_bNoCap => bNoCap);
		q_nState	:= SEL(bNoCap, GVL_CM_RSN.AUTO_CHG, GVL_CM_RSN.NO_CAP);
	ELSIF i_stSet.stRemain.bUse AND F_InHhmmWindow(i_nNow := nNow, i_nStart := i_stSet.stRemain.nStart, i_nEnd := i_stSet.stRemain.nEnd) THEN
		// 2) 잔량 방전 (Messis MT_remain_discharge): 잔량 방전량이 있을 때만, 피크 제어량이 더 크면 그 값
		// [14번 수정 2026-11-09: 방전 허용 시간(공통 stDis: 시간·일요일) 밖이면 잔량 방전·피크 제어 모두 0, 상태 DIS_TIME.
		//   원래는 잔량 방전 시간이면 방전 허용 시간을 보지 않고 방전함]
		IF NOT M_DisAllowed(i_stTime := i_stView.stTime) THEN
			q_nState := GVL_CM_RSN.DIS_TIME;
		ELSE
			fRem		:= M_RemainDis(i_stView := i_stView, i_stWin := i_stSet.stRemain, q_bNoCap => bNoCap);
			q_nState	:= SEL(bNoCap, GVL_CM_RSN.REMAIN_DIS, GVL_CM_RSN.NO_CAP);
			IF fRem > 0.0 THEN
				fP := M_NoReverse(i_fReq := MAX(fRem, _fbPeak.q_fCtrl), i_stView := i_stView, q_nRsn => nRsn);
				IF nRsn <> 0 THEN
					q_nState := nRsn;
				END_IF
			END_IF
		END_IF
	ELSIF _fbPeak.q_bNewInterval THEN
		q_nState := GVL_CM_RSN.NEW_INTERVAL;
	ELSIF _fbPeak.q_fCtrl <= 0.0 THEN
		q_nState := GVL_CM_RSN.BELOW_PEAK;
	ELSIF NOT M_DisAllowed(i_stTime := i_stView.stTime) THEN
		q_nState := GVL_CM_RSN.DIS_TIME;
	ELSE
		// 3) 피크 제어 (Messis MT_peak_shaving_mode)
		fP			:= M_NoReverse(i_fReq := _fbPeak.q_fCtrl, i_stView := i_stView, q_nRsn => nRsn);
		q_nState	:= SEL(nRsn <> 0, GVL_CM_RSN.PEAK, nRsn);
	END_IF
END_IF
M_Calc := M_Finish(i_fP := fP);
END_METHOD

METHOD M_CheckSet : WSTRING(63)
M_CheckSet := SUPER^.M_CheckSet();
IF M_CheckSet <> "" THEN
	RETURN;
END_IF
// [결함 13 수정 2026-11-04: 피크 설정이 숫자인지 먼저]
IF NOT (F_RealOk(i_stSet.stPeak.fTarget) AND F_RealOk(i_stSet.stPeak.fBandSens) AND F_RealOk(i_stSet.stPeak.fLoadRatio) AND F_RealOk(i_stSet.stPeak.fMinOut)) THEN
	M_CheckSet := "피크컷: 피크 설정 숫자 아님";
ELSIF i_stSet.stPeak.fTarget < 0.0 OR i_stSet.stPeak.fBandSens < 0.0 OR i_stSet.stPeak.fLoadRatio < 0.0 OR i_stSet.stPeak.fLoadRatio > 1.0 OR i_stSet.stPeak.fMinOut < 0.0 THEN
	M_CheckSet := "피크컷: 목표·감도·부하 비율(0~1)·최소 출력";
ELSIF NOT M_CheckWindow(i_stWin := i_stSet.stAutoChg) THEN
	M_CheckSet := "피크컷: 자동 충전 시간·SOC";
ELSIF NOT M_CheckWindow(i_stWin := i_stSet.stRemain) THEN
	M_CheckSet := "피크컷: 잔량 방전 시간·SOC";
END_IF
END_METHOD

END_FUNCTION_BLOCK

// ---- 20_Module/ControlMode/FB_CmPeakCalc.TcPOU
FUNCTION_BLOCK FB_CmPeakCalc		// 15분 피크 제어량 계산 (Messis ACT_calc_quarter_avg_and_output 이식). 피크컷·통합 모드가 같이 씀
// 구간 = 시계 기준 15분 (매시 00·15·30·45분). 1초마다 수전·부하 평균, 시계 분이 바뀔 때마다 제어량 갱신, 구간 경계에서 0:
//   목표를 넘은 수전 누적 / 남은 분 (10 단위 반올림) × 속도 × (지난 분/15), 가용 출력 · 30초 평균 부하 × fLoadRatio · (30초 평균 부하 − 역송 여유) 상한
// 켜진 모드에서 매 스캔 부름. 모드가 켜질 때 M_Reset
VAR_INPUT
	i_stSet			: ST_CmPeakCalcSet;
	i_fRevMargin	: REAL;				// kW, 역송 방지 여유 (공통 설정 stNoRev.fMargin)
	i_stView		: ST_CtrlModeView;
END_VAR
VAR_OUTPUT
	q_fCtrl			: REAL;		// kW, 피크 제어 방전량 (0 = 제어 안 함). 1분마다 바뀜
	q_bNewInterval	: BOOL;		// 이번 스캔에 새 15분 구간 시작 (1스캔)
	q_nRemainMin	: UINT;		// 구간 남은 분
	q_fExceeded		: REAL;		// 이 구간 목표를 넘은 수전 누적 (kW·분)
	q_fLoad1m		: REAL;		// 직전 1분 평균 부하 (kW, ESS가 없을 때의 수전)
	q_bNoPcc		: BOOL;		// 접속점 계측 무효 (제어량 0, 평균 안 셈)
END_VAR
VAR
	_bInit			: BOOL;
	_nQuarter		: UINT;		// 지금 구간 번호 (시 × 4 + 분 / 15)
	_nPrevSec		: UINT;		// 지난 스캔 시계 초
	_nPrevMin		: UINT;		// 지난 스캔 시계 분
	_nPrevHalf		: UINT;		// 지난 스캔 30초 칸 (0 / 1)
	_n60			: UINT;		// 1분 평균 표본 수
	_n30			: UINT;		// 30초 평균 표본 수
	_fImp1m			: REAL;		// 1분 평균 수전 (kW)
	_fLoad30		: REAL;		// 30초 평균 부하 (kW)
	_fVelocity		: REAL;		// 제어 속도 (F_CmVelocity)
END_VAR
VAR_TEMP
	nQ				: UINT;
	fImp			: REAL;		// 수전 (kW)
	fLoad			: REAL;		// 부하 (kW)
	fCtrl			: REAL;
	nMin			: UINT;		// 구간 시작부터 지난 분
END_VAR

q_bNewInterval := FALSE;
q_bNoPcc := NOT i_stView.stGroup.stPcc.stMeas.stP.bValid;
IF NOT i_stView.stTime.bValid OR i_stSet.fTarget <= 0.0 THEN
	q_fCtrl	:= 0.0;
	_bInit	:= FALSE;
	RETURN;
END_IF

// 1) 구간 시작 (처음 또는 15분 경계). 경계에서는 제어량 0 (Messis: 남은 분 0으로 계산해 0)
nQ := i_stView.stTime.nHour * 4 + i_stView.stTime.nMinute / 15;
IF NOT _bInit OR nQ <> _nQuarter THEN
	q_bNewInterval	:= _bInit;		// 모드가 켜진 첫 스캔은 새 구간으로 보지 않음
	_bInit			:= TRUE;
	_nQuarter		:= nQ;
	_nPrevSec		:= i_stView.stTime.nSecond;
	_nPrevMin		:= i_stView.stTime.nMinute;
	_nPrevHalf		:= i_stView.stTime.nSecond / 30;
	_n60			:= 0;
	_n30			:= 0;
	q_nRemainMin	:= 15 - i_stView.stTime.nMinute MOD 15;
	q_fExceeded		:= 0.0;
	q_fCtrl			:= 0.0;
	_fVelocity		:= F_CmVelocity(i_fH := i_stSet.fTarget);
	RETURN;
END_IF

// 2) 시계의 초가 바뀔 때마다 (분·30초 경계는 시계 값으로 판단: 시계 보정으로 초가 건너뛰어도 밀리지 않음)
IF i_stView.stTime.nSecond <> _nPrevSec THEN
	_nPrevSec := i_stView.stTime.nSecond;
	// 3) 분이 바뀌면 지난 1분 평균으로 제어량 갱신
	IF i_stView.stTime.nMinute <> _nPrevMin THEN
		_nPrevMin		:= i_stView.stTime.nMinute;
		nMin			:= i_stView.stTime.nMinute MOD 15;		// 구간 시작부터 지난 분
		q_nRemainMin	:= 15 - nMin;
		fCtrl			:= 0.0;
		IF _n60 > 0 AND NOT q_bNoPcc THEN
			q_fExceeded := q_fExceeded + (_fImp1m - i_stSet.fTarget);
			IF q_fLoad1m - i_stSet.fTarget > i_stView.stGroup.fPRatedAvail * UINT_TO_REAL(q_nRemainMin / 15) * i_stSet.fBandSens * 0.5 THEN
				fCtrl := MIN(F_CmRoundTens(i_f := q_fExceeded / UINT_TO_REAL(q_nRemainMin)) * _fVelocity * (UINT_TO_REAL(nMin) / 15.0), i_stView.stGroup.fPRatedAvail);
			END_IF
			fCtrl := MIN(fCtrl, _fLoad30 * i_stSet.fLoadRatio);
			fCtrl := MIN(fCtrl, _fLoad30 - i_fRevMargin);
			IF fCtrl <= 1.0 THEN
				fCtrl := 0.0;
			ELSE
				fCtrl := MAX(fCtrl, i_stSet.fMinOut);
			END_IF
			IF _fImp1m - i_stSet.fTarget > 0.0 THEN
				_fVelocity := F_CmVelocity(i_fH := _fImp1m - i_stSet.fTarget);
			END_IF
		END_IF
		q_fCtrl	:= fCtrl;
		_n60	:= 0;			// 다음 1분 평균을 새로 셈 (값은 남김)
	END_IF
	IF i_stView.stTime.nSecond / 30 <> _nPrevHalf THEN
		_nPrevHalf	:= i_stView.stTime.nSecond / 30;
		_n30		:= 0;		// 다음 30초 평균을 새로 셈 (값은 남김)
	END_IF
	// 4) 1초 표본
	IF q_bNoPcc THEN
		q_fCtrl := 0.0;			// 계측 무효: 평균에 넣지 않고 제어 안 함
	ELSE
		_n60	:= _n60 + 1;
		_n30	:= _n30 + 1;
		fImp	:= -i_stView.stGroup.stPcc.stMeas.stP.fValue;			// 수전 + (접속점 P는 공급 +)
		fLoad	:= i_stView.stGroup.fPOut + fImp;							// ESS가 없을 때의 수전
		_fImp1m		:= (_fImp1m * UINT_TO_REAL(_n60 - 1) + fImp) / UINT_TO_REAL(_n60);
		q_fLoad1m	:= (q_fLoad1m * UINT_TO_REAL(_n60 - 1) + fLoad) / UINT_TO_REAL(_n60);
		_fLoad30	:= (_fLoad30 * UINT_TO_REAL(_n30 - 1) + fLoad) / UINT_TO_REAL(_n30);
	END_IF
END_IF

METHOD M_Reset		// 모드가 켜질 때: 구간을 지금부터 다시 셈, 제어량 0
_bInit		:= FALSE;
q_fCtrl		:= 0.0;
q_fExceeded	:= 0.0;
q_fLoad1m	:= 0.0;
_fImp1m		:= 0.0;
_fLoad30	:= 0.0;
END_METHOD

END_FUNCTION_BLOCK

// ---- 20_Module/ControlMode/F_CmVelocity.TcPOU
FUNCTION F_CmVelocity : REAL		// 피크 제어 속도 (Messis getVelocity): 넘는 양이 작을수록 크게. (log10(h + 100) − log10(h)) × 20, h ≤ 0이면 1
VAR_INPUT
	i_fH		: REAL;		// kW, 목표 또는 목표를 넘은 양
END_VAR

IF i_fH <= 0.0 THEN
	F_CmVelocity := 1.0;
ELSE
	F_CmVelocity := (LOG(i_fH + 100.0) - LOG(i_fH)) * 20.0;
END_IF

END_FUNCTION

// ---- 20_Module/ControlMode/F_CmRoundTens.TcPOU
FUNCTION F_CmRoundTens : REAL		// 10 단위 반올림 (Messis roundUpTens)
VAR_INPUT
	i_f			: REAL;
END_VAR

// [결함 13 수정 2026-11-04: NaN·범위 밖이면 REAL_TO_DINT가 FPU 예외 → F_RealToDint (NaN은 0). 원래 DINT_TO_REAL(REAL_TO_DINT(i_f / 10.0)) * 10.0]
F_CmRoundTens := DINT_TO_REAL(F_RealToDint(i_f / 10.0)) * 10.0;

END_FUNCTION

// ---- 20_Module/ControlMode/FB_CmSchedPeak.TcPOU
FUNCTION_BLOCK FB_CmSchedPeak EXTENDS FB_CmTariffBase		// 제어 모드: 통합 = 스케줄 + 피크컷 (Messis SCHEDULE_PS_MODE)
// 우선순위: 잔량 방전 시간 (잔량 방전과 피크 제어 중 큰 값, 방전 허용 시간에만) → 피크 제어가 필요하고 방전 허용 시간이면 (피크 제어량과 시간표 방전 중 큰 값)
//   → 아니면 스케줄 모드와 같음. 시간표는 스케줄 모드와 같은 표, 피크 제어량 계산은 피크컷과 같은 FB_CmPeakCalc
// Messis와 다른 점: 시간표가 충전 칸일 때 피크 제어가 필요하면 피크 제어량만 방전 (Messis는 충전값 크기만큼 방전할 수 있었음)
VAR_INPUT
	i_stTable	: ST_CmScheduleSet;		// 시간표 (스케줄 모드와 같은 GVL_PERSIST.g_stModuleSet.stCmSchedule)
	i_stSet		: ST_CmSchedPeakSet;	// 설정 (GVL_PERSIST.g_stModuleSet.stCmSchedPeak)
END_VAR
VAR_OUTPUT
	q_fPeakCtrl	: REAL;		// 진단: 피크 제어량 (kW, FB_CmPeakCalc)
	q_nRemainMin	: UINT;		// 진단: 15분 구간 남은 분
	q_fExceeded	: REAL;		// 진단: 구간 목표 초과 수전 누적 (kW·분)
	q_fLoad1m	: REAL;		// 진단: 직전 1분 평균 부하 (kW)
END_VAR
VAR
	_fbPeak		: FB_CmPeakCalc;
END_VAR

METHOD M_Enter
VAR_INPUT
	i_stView	: ST_CtrlModeView;
END_VAR
SUPER^.M_Enter(i_stView := i_stView);
_fbPeak.M_Reset();
END_METHOD

METHOD M_Calc : ST_CtrlModeOut
VAR_INPUT
	i_stView	: ST_CtrlModeView;
END_VAR
VAR
	nNow	: UINT;
	fP		: REAL;
	fRem	: REAL;
	nRsn	: UINT;
	bNoCap	: BOOL;
END_VAR
fP := 0.0;
_fbPeak(i_stSet := i_stSet.stPeak, i_fRevMargin := i_stCommon.stNoRev.fMargin, i_stView := i_stView);
q_fPeakCtrl		:= _fbPeak.q_fCtrl;
q_nRemainMin	:= _fbPeak.q_nRemainMin;
q_fExceeded		:= _fbPeak.q_fExceeded;
q_fLoad1m		:= _fbPeak.q_fLoad1m;
IF M_Begin(i_stView := i_stView) THEN
	nNow := F_TimeHhmm(i_stTime := i_stView.stTime);
	M_SchedLookup(i_stTime := i_stView.stTime, iq_stTable := i_stTable);
	IF i_stSet.stRemain.bUse AND F_InHhmmWindow(i_nNow := nNow, i_nStart := i_stSet.stRemain.nStart, i_nEnd := i_stSet.stRemain.nEnd) THEN
		// 1) 잔량 방전
		// [14번 수정 2026-11-09: 방전 허용 시간(공통 stDis: 시간·일요일) 밖이면 잔량 방전·피크 제어 모두 0, 상태 DIS_TIME.
		//   원래는 잔량 방전 시간이면 방전 허용 시간을 보지 않고 방전함]
		IF NOT M_DisAllowed(i_stTime := i_stView.stTime) THEN
			q_nState := GVL_CM_RSN.DIS_TIME;
		ELSE
			fRem		:= M_RemainDis(i_stView := i_stView, i_stWin := i_stSet.stRemain, q_bNoCap => bNoCap);
			q_nState	:= SEL(bNoCap, GVL_CM_RSN.REMAIN_DIS, GVL_CM_RSN.NO_CAP);
			IF fRem > 0.0 THEN
				fP := M_NoReverse(i_fReq := MAX(fRem, _fbPeak.q_fCtrl), i_stView := i_stView, q_nRsn => nRsn);
				IF nRsn <> 0 THEN
					q_nState := nRsn;
				END_IF
			END_IF
		END_IF
	ELSIF _fbPeak.q_fCtrl > 0.0 AND M_DisAllowed(i_stTime := i_stView.stTime) THEN
		// 2) 피크 제어 + 시간표 방전 중 큰 값
		fP			:= M_NoReverse(i_fReq := MAX(_fbPeak.q_fCtrl, MAX(q_fSlotP, 0.0)), i_stView := i_stView, q_nRsn => nRsn);
		q_nState	:= SEL(nRsn <> 0, GVL_CM_RSN.SCHED_PEAK, nRsn);
	ELSE
		// 3) 스케줄만
		fP			:= M_SchedOut(i_stView := i_stView, q_nRsn => nRsn);
		q_nState	:= nRsn;
	END_IF
END_IF
M_Calc := M_Finish(i_fP := fP);
END_METHOD

METHOD M_CheckSet : WSTRING(63)
M_CheckSet := SUPER^.M_CheckSet();
IF M_CheckSet <> "" THEN
	RETURN;
END_IF
M_CheckSet := M_CheckTable(iq_stTable := i_stTable);
IF M_CheckSet <> "" THEN
	RETURN;
END_IF
// [결함 13 수정 2026-11-04: 피크 설정이 숫자인지 먼저]
IF NOT (F_RealOk(i_stSet.stPeak.fTarget) AND F_RealOk(i_stSet.stPeak.fBandSens) AND F_RealOk(i_stSet.stPeak.fLoadRatio) AND F_RealOk(i_stSet.stPeak.fMinOut)) THEN
	M_CheckSet := "통합: 피크 설정 숫자 아님";
ELSIF i_stSet.stPeak.fTarget < 0.0 OR i_stSet.stPeak.fBandSens < 0.0 OR i_stSet.stPeak.fLoadRatio < 0.0 OR i_stSet.stPeak.fLoadRatio > 1.0 OR i_stSet.stPeak.fMinOut < 0.0 THEN
	M_CheckSet := "통합: 목표·감도·부하 비율(0~1)·최소 출력";
ELSIF NOT M_CheckWindow(i_stWin := i_stSet.stRemain) THEN
	M_CheckSet := "통합: 잔량 방전 시간·SOC";
END_IF
END_METHOD

END_FUNCTION_BLOCK

// ---- 20_Module/Common/FB_SocLimit.TcPOU
FUNCTION_BLOCK FB_SocLimit EXTENDS FB_ModuleBase IMPLEMENTS I_BatLimitRule	// SOC 감발·차단·재개 마진 (버스 제한). 기본 SOC 정책 (Auto·Manual 기본 등록)
// 최대 SOC가 상한에 다가가면 충전 한도를, 최소 SOC가 하한에 다가가면 방전 한도를 줄이고, 한계에서 막음
// 막은 뒤에는 SOC가 재개 마진만큼 돌아와야 다시 허용. 다시 허용한 뒤 감발 구간을 지나는 동안 bResume (재개 램프율)
// 출력 한도만 냄 (장비 명령 없음). 한도가 0이면 그 방향 출력 0 = 대기
// nTarget 0 = 모든 버스를 한 인스턴스가 봄 (버스마다 상태를 따로 가짐)
VAR_INPUT
	i_stSet	: ST_SocLimitSet;	// 설정 (MAIN이 GVL_PERSIST.g_stModuleSet 칸을 매 스캔 넘김. 안 넘기면 기본값)
END_VAR
VAR
	(* 버스마다 상태 *)
	_abChgBlock	: ARRAY[1..GVL_PARAM.BAT_COUNT] OF BOOL;	// 충전 막음 (재개 마진 전까지 유지)
	_abDisBlock	: ARRAY[1..GVL_PARAM.BAT_COUNT] OF BOOL;	// 방전 막음
	_abChgResume	: ARRAY[1..GVL_PARAM.BAT_COUNT] OF BOOL;	// 충전 재개 중 (막음이 풀린 뒤 감발 구간)
	_abDisResume	: ARRAY[1..GVL_PARAM.BAT_COUNT] OF BOOL;
	_afChgRatio	: ARRAY[1..GVL_PARAM.BAT_COUNT] OF REAL;	// 진단: 충전 한도 비율 (1 = 안 줄임)
	_afDisRatio	: ARRAY[1..GVL_PARAM.BAT_COUNT] OF REAL;	// 진단: 방전 한도 비율
END_VAR
VAR CONSTANT
	RSN_CHG_DERATE	: UINT := 1;	// 상한 근처 충전 감발
	RSN_CHG_BLOCK	: UINT := 2;	// 상한 충전 막음
	RSN_DIS_DERATE	: UINT := 3;	// 하한 근처 방전 감발
	RSN_DIS_BLOCK	: UINT := 4;	// 하한 방전 막음
	RSN_SOC_INVALID	: UINT := 5;	// SOC 무효
END_VAR

METHOD M_Evaluate : ST_BatLimitOut
VAR_INPUT
	i_stView	: ST_BatLimitView;
END_VAR
VAR
	b	: UINT;
	fChg	: REAL;	// 충전 한도 비율
	fDis	: REAL;	// 방전 한도 비율
END_VAR
b := i_stView.nBatGroup;
IF b < 1 OR b > GVL_PARAM.BAT_COUNT THEN
	RETURN;
END_IF
// SOC 무효: 상태를 풀고, 설정이면 충·방전 모두 막음
IF NOT i_stView.stSocMax.bValid OR NOT i_stView.stSocMin.bValid THEN
	_abChgBlock[b]	:= FALSE;
	_abDisBlock[b]	:= FALSE;
	_abChgResume[b]	:= FALSE;
	_abDisResume[b]	:= FALSE;
	_afChgRatio[b]	:= 1.0;
	_afDisRatio[b]	:= 1.0;
	IF i_stSet.bBlockOnInvalid THEN
		M_Evaluate.stP.bActive	:= TRUE;
		M_Evaluate.stP.fMax	:= 0.0;
		M_Evaluate.stP.fMin	:= 0.0;
		M_Evaluate.stP.nReason	:= RSN_SOC_INVALID;
		_afChgRatio[b]	:= 0.0;
		_afDisRatio[b]	:= 0.0;
	END_IF
	RETURN;
END_IF

// 충전: 최대 SOC 기준
IF i_stView.stSocMax.fValue >= i_stSet.fSocMax THEN
	_abChgBlock[b]	:= TRUE;
	_abChgResume[b]	:= FALSE;
ELSIF _abChgBlock[b] AND i_stView.stSocMax.fValue <= i_stSet.fSocMax - i_stSet.fResumeMargin THEN
	_abChgBlock[b]	:= FALSE;
	_abChgResume[b]	:= TRUE;
END_IF
fChg := 0.0;
IF NOT _abChgBlock[b] THEN
	fChg := F_SocDerate(i_fSoc := i_stView.stSocMax.fValue, i_fLimit := i_stSet.fSocMax, i_fBand := i_stSet.fBand, i_bUpper := TRUE);
END_IF
IF fChg >= 1.0 THEN
	_abChgResume[b] := FALSE;
END_IF

// 방전: 최소 SOC 기준
IF i_stView.stSocMin.fValue <= i_stSet.fSocMin THEN
	_abDisBlock[b]	:= TRUE;
	_abDisResume[b]	:= FALSE;
ELSIF _abDisBlock[b] AND i_stView.stSocMin.fValue >= i_stSet.fSocMin + i_stSet.fResumeMargin THEN
	_abDisBlock[b]	:= FALSE;
	_abDisResume[b]	:= TRUE;
END_IF
fDis := 0.0;
IF NOT _abDisBlock[b] THEN
	fDis := F_SocDerate(i_fSoc := i_stView.stSocMin.fValue, i_fLimit := i_stSet.fSocMin, i_fBand := i_stSet.fBand, i_bUpper := FALSE);
END_IF
IF fDis >= 1.0 THEN
	_abDisResume[b] := FALSE;
END_IF

_afChgRatio[b]	:= fChg;
_afDisRatio[b]	:= fDis;
M_Evaluate.bResume := _abChgResume[b] OR _abDisResume[b];
IF fChg < 1.0 OR fDis < 1.0 THEN
	M_Evaluate.stP.bActive	:= TRUE;
	M_Evaluate.stP.fMax	:= MAX(i_stView.fPDisMax, 0.0) * fDis;
	M_Evaluate.stP.fMin	:= -MAX(i_stView.fPChgMax, 0.0) * fChg;
	// 이유: 막음이 감발보다 먼저 (한 줄 제한이라 상·하한이 같은 이유를 가짐)
	IF _abDisBlock[b] THEN
		M_Evaluate.stP.nReason := RSN_DIS_BLOCK;
	ELSIF _abChgBlock[b] THEN
		M_Evaluate.stP.nReason := RSN_CHG_BLOCK;
	ELSIF fDis < 1.0 THEN
		M_Evaluate.stP.nReason := RSN_DIS_DERATE;
	ELSE
		M_Evaluate.stP.nReason := RSN_CHG_DERATE;
	END_IF
END_IF
END_METHOD

METHOD M_ReasonText : WSTRING(63)
VAR_INPUT
	i_nReason	: UINT;
END_VAR
CASE i_nReason OF
	RSN_CHG_DERATE:	M_ReasonText := "SOC 상한 근처 충전 감발";
	RSN_CHG_BLOCK:	M_ReasonText := "SOC 상한 충전 막음";
	RSN_DIS_DERATE:	M_ReasonText := "SOC 하한 근처 방전 감발";
	RSN_DIS_BLOCK:	M_ReasonText := "SOC 하한 방전 막음";
	RSN_SOC_INVALID:	M_ReasonText := "SOC 무효";
ELSE
	M_ReasonText := WCONCAT("이유 ", TO_WSTRING(i_nReason));
END_CASE
END_METHOD

METHOD M_CheckSet : WSTRING(63)		// 설정 점검: SOC 상·하한, 감발 폭, 재개 마진
// [9-21 수정 2026-11-04: 검사 규칙을 F_SocLimitSetErr로 옮김 (EMS config 반영 FB_EmsConfigApply와 같은 규칙을 씀). 원래:
//   M_CheckSet := "";
//   IF NOT (F_RealOk(i_stSet.fSocMin) AND F_RealOk(i_stSet.fSocMax) AND F_RealOk(i_stSet.fBand) AND F_RealOk(i_stSet.fResumeMargin)) THEN	// [결함 13 수정 2026-11-04]
//   	M_CheckSet := "SOC 설정 숫자 아님";
//   ELSIF i_stSet.fSocMin < 0.0 OR i_stSet.fSocMax > 100.0 OR i_stSet.fSocMin >= i_stSet.fSocMax THEN
//   	M_CheckSet := "SOC 상·하한 (0 ≤ 하한 < 상한 ≤ 100)";
//   ELSIF i_stSet.fBand < 0.0 OR i_stSet.fSocMin + i_stSet.fBand > i_stSet.fSocMax - i_stSet.fBand THEN
//   	M_CheckSet := "감발 폭 fBand (0 이상, 상·하한 사이)";
//   ELSIF i_stSet.fResumeMargin < 0.0 OR i_stSet.fSocMin + i_stSet.fResumeMargin >= i_stSet.fSocMax - i_stSet.fResumeMargin THEN
//   	M_CheckSet := "재개 마진 fResumeMargin (0 이상, 상·하한 사이)";
//   END_IF]
M_CheckSet := F_SocLimitSetErr(i_stSet);
END_METHOD

END_FUNCTION_BLOCK

// ---- 20_Module/Common/F_SocDerate.TcPOU
FUNCTION F_SocDerate : REAL	// SOC 감발 비율 (0~1, 상태 없음). 여러 SOC 정책 모듈이 같이 씀
// 상한(i_bUpper = TRUE, 충전 쪽): SOC ≥ 한계면 0, 한계 - 폭 < SOC면 선형으로 줄임, 그 아래는 1
// 하한(i_bUpper = FALSE, 방전 쪽): SOC ≤ 한계면 0, SOC < 한계 + 폭이면 선형으로 줄임, 그 위는 1
VAR_INPUT
	i_fSoc	: REAL;	// %
	i_fLimit	: REAL;	// %, 한계
	i_fBand	: REAL;	// %, 감발 폭. 0 이하면 줄이지 않고 한계에서 0
	i_bUpper	: BOOL;	// TRUE = 상한, FALSE = 하한
END_VAR

IF i_bUpper THEN
	IF i_fSoc >= i_fLimit THEN
		F_SocDerate := 0.0;
	ELSIF i_fBand > 0 AND i_fSoc > i_fLimit - i_fBand THEN
		F_SocDerate := (i_fLimit - i_fSoc) / i_fBand;
	ELSE
		F_SocDerate := 1.0;
	END_IF
ELSE
	IF i_fSoc <= i_fLimit THEN
		F_SocDerate := 0.0;
	ELSIF i_fBand > 0 AND i_fSoc < i_fLimit + i_fBand THEN
		F_SocDerate := (i_fSoc - i_fLimit) / i_fBand;
	ELSE
		F_SocDerate := 1.0;
	END_IF
END_IF

END_FUNCTION

// ---- 20_Module/Common/FB_UnitLimit.TcPOU
FUNCTION_BLOCK FB_UnitLimit EXTENDS FB_ModuleBase IMPLEMENTS I_UnitLimitRule	// 사용자 한도: 유닛마다 운전원이 정한 P·Q 상·하한 (kW·kvar). 정격·Derate와 겹쳐 좁은 쪽 (코어 FB_EquipmentLimits)
// 등록: g_aipUnitRule 한 칸, g_astUnitRuleReg nTarget 0 (전체 유닛, 유닛마다 설정을 따로 봄), bAuto·bManual로 적용 모드
// 출력 제한 이유: 유닛 한도 UnitRule + 이 모듈 ID, 이유 "사용자 한도"
VAR_INPUT
	i_stSet		: ST_UnitLimitSet;	// 유닛마다 한도 (MAIN A_PassModuleSet이 g_stModuleSet 칸을 넘김. 안 넘기면 모두 끔)
END_VAR
VAR CONSTANT
	RSN_USER	: UINT := 1;		// 사용자 한도
END_VAR

METHOD M_Evaluate : ST_LimitOut
VAR_INPUT
	i_stView	: ST_UnitLimitView;
END_VAR
VAR
	u	: UINT;
END_VAR
u := i_stView.nUnit;
IF u < 1 OR u > GVL_PARAM.UNIT_COUNT THEN
	RETURN;
END_IF
IF i_stSet.astUnit[u].bPEnable THEN
	M_Evaluate.stP.bActive	:= TRUE;
	M_Evaluate.stP.fMax		:= i_stSet.astUnit[u].fPMax;
	M_Evaluate.stP.fMin		:= i_stSet.astUnit[u].fPMin;
	M_Evaluate.stP.nReason	:= RSN_USER;
END_IF
IF i_stSet.astUnit[u].bQEnable THEN
	M_Evaluate.stQ.bActive	:= TRUE;
	M_Evaluate.stQ.fMax		:= i_stSet.astUnit[u].fQMax;
	M_Evaluate.stQ.fMin		:= i_stSet.astUnit[u].fQMin;
	M_Evaluate.stQ.nReason	:= RSN_USER;
END_IF
END_METHOD

METHOD M_ReasonText : WSTRING(63)
VAR_INPUT
	i_nReason	: UINT;
END_VAR
IF i_nReason = RSN_USER THEN
	M_ReasonText := "사용자 한도";
ELSE
	M_ReasonText := WCONCAT("이유 ", TO_WSTRING(i_nReason));
END_IF
END_METHOD

METHOD M_CheckSet : WSTRING(63)		// 설정 점검: 켠 한도는 상한 ≥ 0 ≥ 하한
VAR
	u	: UINT;
END_VAR
M_CheckSet := "";
FOR u := 1 TO GVL_PARAM.UNIT_COUNT DO
	IF NOT (F_RealOk(i_stSet.astUnit[u].fPMax) AND F_RealOk(i_stSet.astUnit[u].fPMin) AND F_RealOk(i_stSet.astUnit[u].fQMax) AND F_RealOk(i_stSet.astUnit[u].fQMin)) THEN	// [결함 13 수정 2026-11-04]
		M_CheckSet := F_TxtNum("한도 숫자 아님: 유닛 ", u);
		RETURN;
	END_IF
	IF i_stSet.astUnit[u].bPEnable AND (i_stSet.astUnit[u].fPMax < 0.0 OR i_stSet.astUnit[u].fPMin > 0.0) THEN
		M_CheckSet := F_TxtNum("P 한도 상한 < 0 또는 하한 > 0: 유닛 ", u);
		RETURN;
	END_IF
	IF i_stSet.astUnit[u].bQEnable AND (i_stSet.astUnit[u].fQMax < 0.0 OR i_stSet.astUnit[u].fQMin > 0.0) THEN
		M_CheckSet := F_TxtNum("Q 한도 상한 < 0 또는 하한 > 0: 유닛 ", u);
		RETURN;
	END_IF
END_FOR
END_METHOD

END_FUNCTION_BLOCK

// ---- 20_Module/Standard/FB_ProtPcsFault.TcPOU
FUNCTION_BLOCK FB_ProtPcsFault EXTENDS FB_ModuleBase IMPLEMENTS I_ProtectionRule		// 표준 보호: PCS 고장 (범위 Unit): 통신이 있고 PCS가 고장을 알림. 기본 등록. 빼면 이 보호 없음. 현장마다 다르면 복사해 이름을 바꿔 그 칸에 대신 등록
VAR
END_VAR

METHOD M_Evaluate : BOOL		// 범위가 맞지 않게 등록되면 FALSE (보호 안 걸림)
VAR_INPUT
	i_stView	: ST_ProtView;
END_VAR
M_Evaluate := i_stView.eScope = E_ProtScope.Unit AND i_stView.bInstalled AND i_stView.stUnit.bComm AND i_stView.stUnit.bFault;
END_METHOD

END_FUNCTION_BLOCK

// ---- 20_Module/Standard/FB_ProtPcsComm.TcPOU
FUNCTION_BLOCK FB_ProtPcsComm EXTENDS FB_ModuleBase IMPLEMENTS I_ProtectionRule		// 표준 보호: PCS 통신 끊김 (범위 Unit). 기본 등록. 빼면 이 보호 없음. 현장마다 다르면 복사해 이름을 바꿔 그 칸에 대신 등록
VAR
END_VAR

METHOD M_Evaluate : BOOL		// 범위가 맞지 않게 등록되면 FALSE (보호 안 걸림)
VAR_INPUT
	i_stView	: ST_ProtView;
END_VAR
M_Evaluate := i_stView.eScope = E_ProtScope.Unit AND i_stView.bInstalled AND NOT i_stView.stUnit.bComm;
END_METHOD

END_FUNCTION_BLOCK

// ---- 20_Module/Standard/FB_ProtBmsFault.TcPOU
FUNCTION_BLOCK FB_ProtBmsFault EXTENDS FB_ModuleBase IMPLEMENTS I_ProtectionRule		// 표준 보호: BMS 고장 (범위 Bms): 통신이 있고 BMS가 고장을 알림. 기본 등록. 빼면 이 보호 없음. 현장마다 다르면 복사해 이름을 바꿔 그 칸에 대신 등록
VAR
END_VAR

METHOD M_Evaluate : BOOL		// 범위가 맞지 않게 등록되면 FALSE (보호 안 걸림)
VAR_INPUT
	i_stView	: ST_ProtView;
END_VAR
M_Evaluate := i_stView.eScope = E_ProtScope.Bms AND i_stView.bInstalled AND i_stView.stBms.bComm AND i_stView.stBms.bFault;
END_METHOD

END_FUNCTION_BLOCK

// ---- 20_Module/Standard/FB_ProtBmsComm.TcPOU
FUNCTION_BLOCK FB_ProtBmsComm EXTENDS FB_ModuleBase IMPLEMENTS I_ProtectionRule		// 표준 보호: BMS 통신 끊김 (범위 Bms). 기본 등록. 빼면 이 보호 없음. 현장마다 다르면 복사해 이름을 바꿔 그 칸에 대신 등록
VAR
END_VAR

METHOD M_Evaluate : BOOL		// 범위가 맞지 않게 등록되면 FALSE (보호 안 걸림)
VAR_INPUT
	i_stView	: ST_ProtView;
END_VAR
M_Evaluate := i_stView.eScope = E_ProtScope.Bms AND i_stView.bInstalled AND NOT i_stView.stBms.bComm;
END_METHOD

END_FUNCTION_BLOCK

// ---- 20_Module/Standard/FB_ProtPccInvalid.TcPOU
FUNCTION_BLOCK FB_ProtPccInvalid EXTENDS FB_ModuleBase IMPLEMENTS I_ProtectionRule		// 표준 보호: 접속점 계측 무효 (범위 Group): 접속점 유효전력 값이 무효. 기본 등록. 빼면 이 보호 없음. 현장마다 다르면 복사해 이름을 바꿔 그 칸에 대신 등록
VAR
END_VAR

METHOD M_Evaluate : BOOL		// 범위가 맞지 않게 등록되면 FALSE (보호 안 걸림)
VAR_INPUT
	i_stView	: ST_ProtView;
END_VAR
// [결함 7 수정 2026-11-03: 접속점이 없는 그룹(nPccPoint 0)은 판단 안 함. 원래 M_Evaluate := i_stView.eScope = E_ProtScope.Group AND NOT i_stView.stPcc.stMeas.stP.bValid;]
M_Evaluate := i_stView.eScope = E_ProtScope.Group AND NOT i_stView.stPcc.bNoPoint AND NOT i_stView.stPcc.stMeas.stP.bValid;
END_METHOD

END_FUNCTION_BLOCK

// ---- 20_Module/Standard/FB_ProtRespStd.TcPOU
FUNCTION_BLOCK FB_ProtRespStd EXTENDS FB_ModuleBase IMPLEMENTS I_ProtResponse		// 표준 보호 대응 (기본 등록: GVL_SITE.g_aipResp 칸마다 같은 인스턴스): 칸 설정(ST_ProtCfg)의 조치를 범위 안 유닛·BMS에 한 단계로 요청
// 유닛: 범위에 드는 유닛 중 그 운전 모드에 조치를 거는 것(bAuto·bManual)만. 모드 조치(ToManual)는 bAuto 항목이면 범위 안 유닛 전부
// BMS: Bms·BatGroup 범위는 그 버스에 조치를 받는 유닛이 있을 때 (버스에 유닛이 없으면 그대로). Unit·Group·Site 범위는 조치를 받는 유닛의 배터리 그룹 BMS 전부
// 현장 대응이 다르면 이 FB를 복사해 이름을 바꿔 그 칸에 대신 등록. 상태가 없어 인스턴스 하나를 모든 칸에 같이 등록함

METHOD M_Respond		// 칸 설정(stProt)의 조치를 걸렸을 때만 요청
// 코어가 매 스캔 범위 안 대상마다 부름 (조건이 없을 때도: 단계 대응의 타이머·상태를 풀 수 있게). 대상 번호가 0으로 등록되면 대상마다 상태를 따로 둠
VAR_INPUT
	i_bActive		: BOOL;			// 보호 조건 있음 (등록 bAuto·bManual 중 하나가 켜져 있고 조건 모듈이 TRUE)
	i_tActive		: TIME;			// 조건이 이어진 시간 (조건 없으면 0)
	i_nTarget		: UINT;			// 대상 번호 (범위는 i_stRule.eScope. Site면 1)
	i_stRule		: ST_RuleCfg;		// 이 칸 설정 (범위·대상·임계값·표준 대응 설정)
END_VAR
VAR_IN_OUT CONSTANT
	iq_astUnit		: ARRAY[1..GVL_PARAM.UNIT_COUNT] OF ST_UnitState;	// 장비 상태 (이번 스캔 스냅샷, 읽기 전용)
	iq_astBms		: ARRAY[1..GVL_PARAM.BMS_COUNT] OF ST_BatState;
	iq_astUnitCfg	: ARRAY[1..GVL_PARAM.UNIT_COUNT] OF ST_UnitCfg;		// 소속 (제어 그룹·배터리 그룹)
	iq_astBmsCfg	: ARRAY[1..GVL_PARAM.BMS_COUNT] OF ST_BmsCfg;
	iq_aeOpMode		: ARRAY[1..GVL_PARAM.UNIT_COUNT] OF E_OpMode;		// 실제 운전 모드
END_VAR
VAR_IN_OUT
	iq_stReq		: ST_ProtReq;		// 요청 (코어가 비워서 넘김)
END_VAR
VAR
	u			: UINT;
	m			: UINT;
	nBus		: UINT;		// Bms·BatGroup 범위의 배터리 그룹
	nBusUnits	: UINT;		// 그 버스의 유닛 수
	bBusTakes	: BOOL;		// 그 버스에 조치를 받는 유닛이 있음
	bIn			: BOOL;
	bManual		: BOOL;
	bTakes		: BOOL;
	stCfg		: ST_ProtCfg;
END_VAR
IF NOT i_bActive THEN
	RETURN;
END_IF
stCfg := i_stRule.stProt;
nBus := 0;
IF i_stRule.eScope = E_ProtScope.Bms AND i_nTarget >= 1 AND i_nTarget <= GVL_PARAM.BMS_COUNT THEN
	nBus := iq_astBmsCfg[i_nTarget].nBatGroup;
ELSIF i_stRule.eScope = E_ProtScope.BatGroup THEN
	nBus := i_nTarget;
END_IF
(* 1) 유닛 *)
nBusUnits := 0;
bBusTakes := FALSE;
FOR u := 1 TO GVL_PARAM.UNIT_COUNT DO
	CASE i_stRule.eScope OF
		E_ProtScope.Unit:					bIn := u = i_nTarget;
		E_ProtScope.Bms, E_ProtScope.BatGroup:	bIn := nBus <> 0 AND iq_astUnitCfg[u].nBatGroup = nBus;
		E_ProtScope.Group:					bIn := iq_astUnitCfg[u].nGroup = i_nTarget;
		E_ProtScope.Site:					bIn := TRUE;
	ELSE
		bIn := FALSE;
	END_CASE
	IF bIn THEN
		bManual	:= iq_aeOpMode[u] = E_OpMode.Manual;
		bTakes	:= F_ModeApplies(stCfg.bAuto, stCfg.bManual, BOOL_TO_UINT(NOT bManual), BOOL_TO_UINT(bManual));
		nBusUnits := nBusUnits + 1;
		bBusTakes := bBusTakes OR bTakes;
		// 모드 조치: Auto 유닛에 거는 항목이면 실제 모드와 관계없이 (이미 Manual이어도 Auto 재요청을 막음)
		IF stCfg.bAuto AND stCfg.eModeAction = E_ModeAction.ToManual THEN
			iq_stReq.abToManual[u] := TRUE;
		END_IF
		IF bTakes THEN
			iq_stReq.aePcs[u]	:= stCfg.ePcsAction;
			iq_stReq.afPPct[u]	:= stCfg.fPPct;
			iq_stReq.afQPct[u]	:= stCfg.fQPct;
			// 유닛·제어 그룹·사이트 범위: 그 유닛 배터리 그룹의 BMS 전부
			IF stCfg.eBatAction <> E_BatAction.None AND nBus = 0 AND iq_astUnitCfg[u].nBatGroup <> 0 THEN
				FOR m := 1 TO GVL_PARAM.BMS_COUNT DO
					IF iq_astBmsCfg[m].nBatGroup = iq_astUnitCfg[u].nBatGroup THEN
						iq_stReq.aeBat[m] := stCfg.eBatAction;
					END_IF
				END_FOR
			END_IF
		END_IF
	END_IF
END_FOR
(* 2) Bms·BatGroup 범위의 배터리 조치: 버스에 조치를 받는 유닛이 있을 때 (버스에 유닛이 없으면 그대로) *)
IF nBus <> 0 AND stCfg.eBatAction <> E_BatAction.None AND (bBusTakes OR nBusUnits = 0) THEN
	FOR m := 1 TO GVL_PARAM.BMS_COUNT DO
		IF (i_stRule.eScope = E_ProtScope.Bms AND m = i_nTarget) OR (i_stRule.eScope = E_ProtScope.BatGroup AND iq_astBmsCfg[m].nBatGroup = nBus) THEN
			iq_stReq.aeBat[m] := stCfg.eBatAction;
		END_IF
	END_FOR
END_IF
END_METHOD

END_FUNCTION_BLOCK

// ---- 20_Module/Common/FB_RuleValue.TcPOU
FUNCTION_BLOCK FB_RuleValue EXTENDS FB_ModuleBase IMPLEMENTS I_ProtectionRule, I_OutputRule		// 아날로그 값 하나 ↔ 임계값 (온도·습도 등). 임계값은 등록 설정(fThreshold)에서 받음
VAR_INPUT
	i_ipAux			: I_AuxDevice;		// 읽을 보조 장비 (선언 때 지정)
	i_nPoint		: UINT;				// 아날로그 입력 점 번호
	i_stSet			: ST_RuleValueSet;	// 설정: 이하·이상, 해소 폭, 통신 끊김 시 조건 (MAIN이 GVL_PERSIST.g_stModuleSet 칸을 매 스캔 넘김. 안 넘기면 기본값)
END_VAR
VAR
	_bProtCond		: BOOL;				// 보호 규칙 판단 상태 (히스테리시스)
	_bOutCond		: BOOL;				// 출력 규칙 판단 상태 (히스테리시스)
END_VAR

METHOD M_Evaluate : BOOL		// 보호 규칙으로 판단 (보호용 상태 _bProtCond. 값 하나라 대상과 관계없음)
VAR_INPUT
	i_stView	: ST_ProtView;
END_VAR
M_Evaluate := M_Judge(i_fThreshold := i_stView.fThreshold, iq_bCond := _bProtCond);
END_METHOD

METHOD M_Check : BOOL		// 출력 규칙으로 판단 (출력용 상태 _bOutCond. 보호와 같은 인스턴스여도 히스테리시스가 섞이지 않음)
VAR_INPUT
	i_fThreshold	: REAL;
END_VAR
M_Check := M_Judge(i_fThreshold := i_fThreshold, iq_bCond := _bOutCond);
END_METHOD

METHOD PRIVATE M_Judge : BOOL		// 임계값·히스테리시스 판단. 상태는 부르는 쪽 것을 씀
VAR_INPUT
	i_fThreshold	: REAL;
END_VAR
VAR_IN_OUT
	iq_bCond		: BOOL;			// 이 판단의 히스테리시스 상태 (보호용·출력용 따로)
END_VAR
VAR
	stValue			: ST_Val;
END_VAR
IF i_ipAux = 0 THEN
	iq_bCond := FALSE;
ELSE
	stValue := i_ipAux.M_GetValue(i_nPoint);
	IF NOT i_ipAux.Comm OR NOT stValue.bValid THEN
		iq_bCond := i_stSet.bOnCommLoss;
	ELSIF NOT i_stSet.bBelow THEN
		IF stValue.fValue >= i_fThreshold THEN
			iq_bCond := TRUE;
		ELSIF stValue.fValue < i_fThreshold - i_stSet.fHyst THEN
			iq_bCond := FALSE;
		END_IF
	ELSE
		IF stValue.fValue <= i_fThreshold THEN
			iq_bCond := TRUE;
		ELSIF stValue.fValue > i_fThreshold + i_stSet.fHyst THEN
			iq_bCond := FALSE;
		END_IF
	END_IF
END_IF
M_Judge := iq_bCond;
END_METHOD

METHOD M_CheckSet : WSTRING(63)		// 설정 점검: 해소 폭 (FB_RuleBit은 점검할 값 없음)
M_CheckSet := "";
IF NOT F_RealOk(i_stSet.fHyst) THEN	// [결함 13 수정 2026-11-04]
	M_CheckSet := "해소 폭 fHyst 숫자 아님";
ELSIF i_stSet.fHyst < 0.0 THEN
	M_CheckSet := "해소 폭 fHyst 음수";
END_IF
END_METHOD

END_FUNCTION_BLOCK

// ---- 20_Module/Common/FB_BreakerCtrl.TcPOU
FUNCTION_BLOCK FB_BreakerCtrl EXTENDS FB_ModuleBase IMPLEMENTS I_OutputRule, I_ProtectionRule	// 차단기(VCB) 운전원 투입·개방: 지령 → 코일 펄스(DO) → 상태 접점 확인 → 실패 감시
// 출력: 출력 규칙 칸 두 개에 같은 인스턴스를 등록하고 g_astOutputCfg의 fThreshold로 코일을 고름 (1 = 투입 코일, 2 = 개방 코일). 장비·점은 그 칸의 nAux·nPoint, 지연 0·유지 끔
// 실패 감시: 보호 규칙 칸에도 같은 인스턴스를 등록 (g_astRuleCfg 조치 None이면 알람만). 조건 = 투입 실패 또는 개방 실패 (다음 성공 조작 또는 i_bResetFail로 풀림)
// 지령: HMI가 i_bCloseCmd·i_bOpenCmd를 켬 (상승 에지 1번에 1회). 같이 오면 개방이 이김. 투입은 상태 접점이 정상이고 개방 상태일 때만, 개방은 언제나 (조작 중이어도 끼어듦)
// 보호 트립 같은 자동 개방은 다른 출력 규칙(FB_RuleBit 등)을 같은 개방 코일 점에 등록 (같은 점은 OR)
// 스캔마다 한 번만 갱신 (보호 규칙·출력 규칙으로 여러 번 불려도 첫 호출에서만)
VAR_INPUT
	i_ipAux			: I_AuxDevice;		// 상태 접점을 읽을 보조 장비 (선언 때 지정)
	i_nClosedPoint	: UINT;				// 디지털 입력 점: TRUE = 투입 상태
	i_stSet			: ST_BreakerSet;	// 펄스 폭·확인 시간 (MAIN A_PassModuleSet이 g_stModuleSet 칸을 넘김. 안 넘기면 기본값)
	i_bCloseCmd		: BOOL;				// 투입 지령 (HMI, 상승 에지)
	i_bOpenCmd		: BOOL;				// 개방 지령 (HMI, 상승 에지)
	i_bResetFail	: BOOL;				// 실패 표시 풀기 (HMI, 상승 에지)
END_VAR
VAR_OUTPUT
	q_bClosed		: BOOL;		// 투입 상태 (상태 접점, 마지막으로 읽은 값)
	q_bStateValid	: BOOL;		// 상태 접점을 읽을 수 있음 (보조 장비 통신 정상)
	q_bClosePulse	: BOOL;		// 투입 코일 출력 중
	q_bOpenPulse	: BOOL;		// 개방 코일 출력 중
	q_bBusy			: BOOL;		// 조작 확인 중
	q_bCloseFail	: BOOL;		// 투입 실패 (확인 시간 안에 투입 상태가 안 됨)
	q_bOpenFail		: BOOL;		// 개방 실패
END_VAR
VAR
	_rtClose		: R_TRIG;
	_rtOpen			: R_TRIG;
	_rtReset		: R_TRIG;
	_tonPulse		: TON;
	_tonConfirm		: TON;
	_nOp			: INT;		// 진행 중인 조작 (OP_NONE / OP_CLOSE / OP_OPEN)
	_fbTask			: GETCURTASKINDEX;
	_nLastCycle		: UDINT;
	_bRan			: BOOL;
END_VAR
VAR CONSTANT
	OP_NONE			: INT := 0;
	OP_CLOSE		: INT := 1;
	OP_OPEN			: INT := 2;
	COIL_CLOSE		: REAL := 1.0;	// 출력 규칙 fThreshold: 투입 코일
	COIL_OPEN		: REAL := 2.0;	// 개방 코일
	RSN_CLOSE_FAIL	: UINT := 1;
	RSN_OPEN_FAIL	: UINT := 2;
END_VAR

METHOD PRIVATE M_Update		// 스캔마다 한 번: 상태 읽기 → 지령 → 펄스 → 확인
VAR
	nCycle	: UDINT;
	bNew	: BOOL;
END_VAR
_fbTask();
nCycle := TwinCAT_SystemInfoVarList._TaskInfo[_fbTask.index].CycleCount;
IF _bRan AND nCycle = _nLastCycle THEN
	RETURN;		// 이번 스캔은 이미 갱신함
END_IF
_bRan		:= TRUE;
_nLastCycle	:= nCycle;

// 상태 접점
q_bStateValid := FALSE;
IF i_ipAux <> 0 THEN
	q_bStateValid := i_ipAux.Comm;
	IF q_bStateValid THEN
		q_bClosed := i_ipAux.M_GetBit(i_nClosedPoint);
	END_IF
END_IF

// 지령 (개방이 이김. 투입은 상태를 알고 개방 상태일 때만, 진행 중인 조작이 없을 때만)
_rtClose(CLK := i_bCloseCmd);
_rtOpen(CLK := i_bOpenCmd);
_rtReset(CLK := i_bResetFail);
IF _rtReset.Q THEN
	q_bCloseFail	:= FALSE;
	q_bOpenFail		:= FALSE;
END_IF
bNew := FALSE;
IF _rtOpen.Q AND NOT (q_bStateValid AND NOT q_bClosed) THEN
	_nOp	:= OP_OPEN;
	bNew	:= TRUE;
ELSIF _rtClose.Q AND _nOp = OP_NONE AND q_bStateValid AND NOT q_bClosed THEN
	_nOp	:= OP_CLOSE;
	bNew	:= TRUE;
END_IF
IF bNew THEN
	_tonPulse(IN := FALSE);
	_tonConfirm(IN := FALSE);
END_IF

// 펄스·확인
_tonPulse(IN := _nOp <> OP_NONE, PT := i_stSet.tPulse);
_tonConfirm(IN := _nOp <> OP_NONE, PT := i_stSet.tConfirm);
q_bClosePulse	:= _nOp = OP_CLOSE AND NOT _tonPulse.Q;
q_bOpenPulse	:= _nOp = OP_OPEN AND NOT _tonPulse.Q;
IF _nOp = OP_CLOSE THEN
	IF q_bStateValid AND q_bClosed THEN
		_nOp			:= OP_NONE;
		q_bCloseFail	:= FALSE;
	ELSIF _tonConfirm.Q THEN
		_nOp			:= OP_NONE;
		q_bCloseFail	:= TRUE;
	END_IF
ELSIF _nOp = OP_OPEN THEN
	IF q_bStateValid AND NOT q_bClosed THEN
		_nOp			:= OP_NONE;
		q_bOpenFail		:= FALSE;
	ELSIF _tonConfirm.Q THEN
		_nOp			:= OP_NONE;
		q_bOpenFail		:= TRUE;
	END_IF
END_IF
q_bBusy := _nOp <> OP_NONE;
END_METHOD

METHOD M_Check : BOOL		// 출력 규칙: fThreshold 1 = 투입 코일, 2 = 개방 코일
VAR_INPUT
	i_fThreshold	: REAL;
END_VAR
M_Update();
IF i_fThreshold = COIL_CLOSE THEN
	M_Check := q_bClosePulse;
ELSIF i_fThreshold = COIL_OPEN THEN
	M_Check := q_bOpenPulse;
ELSE
	M_Check := FALSE;
END_IF
END_METHOD

METHOD M_Evaluate : BOOL		// 보호 규칙: 투입 실패 또는 개방 실패
VAR_INPUT
	i_stView	: ST_ProtView;	// 안 씀 (차단기 하나)
END_VAR
M_Update();
M_Evaluate := q_bCloseFail OR q_bOpenFail;
END_METHOD

METHOD M_ReasonText : WSTRING(63)
VAR_INPUT
	i_nReason	: UINT;
END_VAR
CASE i_nReason OF
	RSN_CLOSE_FAIL:	M_ReasonText := "차단기 투입 실패";
	RSN_OPEN_FAIL:	M_ReasonText := "차단기 개방 실패";
ELSE
	M_ReasonText := WCONCAT("이유 ", TO_WSTRING(i_nReason));
END_CASE
END_METHOD

METHOD M_CheckSet : WSTRING(63)		// 설정 점검: 펄스 폭, 확인 시간
M_CheckSet := "";
IF i_stSet.tPulse = T#0S THEN
	M_CheckSet := "펄스 폭 tPulse 0";
ELSIF i_stSet.tConfirm < i_stSet.tPulse THEN
	M_CheckSet := "확인 시간 tConfirm이 펄스 폭보다 짧음";
END_IF
END_METHOD

END_FUNCTION_BLOCK

// ---- 20_Module/Virtual/FB_BmsSim.TcPOU
FUNCTION_BLOCK FB_BmsSim EXTENDS FB_DeviceBase IMPLEMENTS I_Bms		// 가상 배터리 (시험용)
VAR_INPUT
	i_fPDc			: REAL;				// kW, 배터리에서 나가는 전력 (방전 +). PRG_SimLink가 넣음
	i_fSocInit		: REAL := 50.0;		// %
	i_fCapacity		: REAL := 4000.0;	// kWh
	i_fPLimit		: REAL := 2000.0;	// kW, 충·방전 한도
	i_bForceFault	: BOOL;				// 시험: 배터리 고장
	i_bForceSysStop	: BOOL;				// 시험: 시스템 정지
	i_bForceCommLoss	: BOOL;			// 시험: 응답 안 함. i_tCommTimeout 뒤 통신 이상
	i_bIgnoreCmd	: BOOL;				// 시험: 상태 명령을 접수하되 접촉기는 바꾸지 않음
	i_bDisableAutoOpen : BOOL;		// 시험: 고장·시스템 정지 때 자동 개방 안 함 (명령에 의한 개방은 별도)
END_VAR
VAR
	_bInit			: BOOL;
	_bClosed		: BOOL;
	_fSoc			: REAL;
	_stBat			: ST_BatState;
END_VAR

PROPERTY BatState : ST_BatState
GET
BatState := _stBat;
END_GET
END_PROPERTY

METHOD M_Cycle
VAR
	fDtHour		: REAL;
END_VAR
IF M_IsReadTime() AND NOT i_bForceCommLoss THEN		// 시험: 통신 끊김이면 응답 안 함
	M_MarkAlive();
END_IF
M_UpdateComm();

IF NOT _bInit THEN
	_fSoc	:= i_fSocInit;
	_bInit	:= TRUE;
END_IF

// 고장·시스템 정지면 접촉기 개방 (시험 입력으로 자동 개방만 끌 수 있음)
IF (i_bForceFault OR i_bForceSysStop) AND NOT i_bDisableAutoOpen THEN
	_bClosed := FALSE;
END_IF

// SOC 적분 (접촉기 투입 중일 때만)
IF _bClosed AND i_fCapacity > 0 THEN
	fDtHour	:= F_CycleSec() / 3600.0;
	_fSoc	:= LIMIT(0.0, _fSoc - i_fPDc * fDtHour / i_fCapacity * 100.0, 100.0);
END_IF

_stBat.bComm			:= _bComm;
_stBat.bContactorClosed	:= _bClosed;
_stBat.bWarn			:= FALSE;
_stBat.bFault			:= i_bForceFault;
_stBat.bSysStop			:= i_bForceSysStop;
_stBat.stSoc.fValue		:= _fSoc;
_stBat.stSoc.bValid		:= TRUE;
_stBat.stSoh.fValue		:= 100.0;
_stBat.stSoh.bValid		:= TRUE;
_stBat.fPChgMax			:= SEL(_fSoc < 100.0, 0.0, i_fPLimit);
_stBat.fPDisMax			:= SEL(_fSoc > 0.0, 0.0, i_fPLimit);
END_METHOD

METHOD M_SetStateCmd : BOOL
VAR_INPUT
	i_stCmd		: ST_BatCmd;
END_VAR
CASE i_stCmd.eCmd OF
	E_BatCmd.Close:
		IF NOT i_bIgnoreCmd AND NOT i_bForceFault AND NOT i_bForceSysStop THEN _bClosed := TRUE; END_IF
	E_BatCmd.Open,
	E_BatCmd.EStop:
		IF NOT i_bIgnoreCmd THEN _bClosed := FALSE; END_IF
	E_BatCmd.Reset:
		;	// 가상 장비는 고장 리셋을 입력(i_bForceFault)으로 함
ELSE
	RETURN;
END_CASE
M_SetStateCmd := TRUE;
END_METHOD

END_FUNCTION_BLOCK

// ---- 20_Module/Ups/FB_UpsChargeRequest.TcPOU
FUNCTION_BLOCK FB_UpsChargeRequest // 요청 번호와 완료 확인 관리
VAR_INPUT
	i_eAction : E_UpsChargeAction;
	i_fValue : REAL;
	i_tTimeout : TIME;
	i_stFeedback : ST_UpsChargeFeedback;
END_VAR
VAR_OUTPUT
	q_stRequest : ST_UpsChargeRequest;
	q_bDone : BOOL;
	q_bError : BOOL;
END_VAR
VAR
	_nSeq : UDINT;
	_ton : TON;
	_bWasPending : BOOL;
END_VAR

_bWasPending := q_stRequest.bValid;
IF i_eAction = E_UpsChargeAction.NoRequest THEN
	q_stRequest.bValid := FALSE;
	q_bDone := FALSE;
	q_bError := FALSE;
ELSE
	IF NOT q_stRequest.bValid AND NOT q_bDone AND NOT q_bError THEN
		_nSeq := F_UpsNextSeq(_nSeq);
		q_stRequest.nSeq := _nSeq;
		q_stRequest.eAction := i_eAction;
		q_stRequest.fValue := i_fValue;
		q_stRequest.bValid := TRUE;
	END_IF
	IF _bWasPending AND i_stFeedback.bValid AND i_stFeedback.nSeq = q_stRequest.nSeq THEN
		q_stRequest.bValid := FALSE;
		q_bDone := i_stFeedback.bConfirmed;
		q_bError := NOT i_stFeedback.bConfirmed;
	END_IF
END_IF
_ton(IN:=q_stRequest.bValid, PT:=i_tTimeout);
IF q_stRequest.bValid AND (_ton.Q OR i_tTimeout = T#0MS) THEN
	q_stRequest.bValid := FALSE;
	q_bError := TRUE;
END_IF

END_FUNCTION_BLOCK

// ---- 20_Module/Ups/FB_UpsChargeSequence.TcPOU
FUNCTION_BLOCK FB_UpsChargeSequence // 충방전 순서에 따른 요청 생성
VAR_INPUT
	i_bEnable : BOOL;
	i_bCancel : BOOL;
	i_bReset : BOOL;
	i_bResetReference : BOOL; // 기준 결과 초기화
	i_eMode : E_UpsChargeMode;
	i_stSet : ST_UpsChargeSet;
	i_stUps : ST_UpsState;
	i_stBms : ST_EsolutionState;
	i_stTime : ST_LocalTime;
	i_stFeedback : ST_UpsChargeFeedback;
END_VAR
VAR_OUTPUT
	q_eStep : E_UpsChargeStep;
	q_eMode : E_UpsChargeMode;
	q_stRequest : ST_UpsChargeRequest;
	q_stActiveSet : ST_UpsChargeSet; // 이번 운전에 고정한 설정
	q_bDone : BOOL; // 정상 완료
	q_bCanceled : BOOL; // 취소 완료
	q_bConflict : BOOL; // 다른 주 운전 시작 충돌
	q_bRecoveryRequired : BOOL; // 현장 상태 확인 필요
	q_nError : UINT; // 1: 설정, 2: 통신/보호, 3: 요청, 4: 모드, 5: 시간 초과
	q_bReferenceValid : BOOL; // 최초 주기적 방전 결과
	q_fReferenceStartVoltageV : REAL;
	q_fReferenceEndVoltageV : REAL;
	q_stReferenceTime : ST_LocalTime;
	q_fStartVoltageV : REAL;
	q_fEndVoltageV : REAL;
	q_stLastTime : ST_LocalTime;
	q_nLastScheduleDate : UDINT;
END_VAR
VAR
	_fbRequest : FB_UpsChargeRequest;
	_eAction : E_UpsChargeAction;
	_bNormal : BOOL;
	_bDataOk : BOOL;
	_bStarted : BOOL;
	_bCanceled : BOOL;
	_bClearRequest : BOOL;
	_bUpsDischargeRequested : BOOL;
	_bDue : BOOL;
	_bEndReached : BOOL;
	_bRestartReached : BOOL;
	_nDate : UDINT;
	_nWeek : UINT;
	_nModeSample : UDINT;
	_tonExtra : TON;
	_tonRest : TON;
	_tonInitial : TON;
	_tonDischarge : TON;
	_tonRun : TON;
	_tonMode : TON;
	_tonAbnormal : TON; // 운전 중 BBC Normal 해제가 이어진 시간
	_bProtTrip : BOOL; // 사고/고장 3~6단계 신호 (동작시퀀스 7쪽)
	_bHardOk : BOOL; // 데이터 유효, 3~6단계·BMS Minor 없음
	_bActive : BOOL; // 운전 단계 (Idle·WaitNormal·Complete·Fault 아님)
	_bWaitStep : BOOL; // 오래 기다리는 단계 (스케줄 대기·휴지)
	_bSafeCancel : BOOL; // 고장 뒤 UPS 방전 취소 요청 중
	_nNewFault : UINT; // 이번 스캔에 생긴 고장 번호
END_VAR

q_bDone := FALSE;
q_bCanceled := FALSE;
IF i_bResetReference AND (q_eStep = E_UpsChargeStep.Idle OR q_eStep = E_UpsChargeStep.WaitSchedule) THEN
	q_bReferenceValid:=FALSE;
END_IF
_eAction := E_UpsChargeAction.NoRequest;
_bClearRequest := FALSE;
_nNewFault := 0;
_bDataOk := i_stUps.bValid AND i_stBms.bValid;
// 동작시퀀스 7쪽 3~6단계: UPS·BMS가 배터리 컨버터 정지·MCCB Trip·컨택터 차단을 하는 상황. 어느 단계에서든 즉시 고장, 자동 재개 없음
// 비상정지(6), BMS Major(3), STATUS2 b12·b13 지락(RCD) 1·2단계(3·4, 명세 v2.50), b14 화재(5), BBC 정지 알람(4), BMS 고장·잠금(5)
_bProtTrip := (i_stUps.bValid AND (i_stUps.bEmergencyStop OR i_stUps.bBmsMajor
		OR (i_stUps.wStatus2 AND 16#7000) <> 0 OR (i_stUps.wBbcAlarm AND 16#0FA8) <> 0))
	OR (i_stBms.bValid AND (i_stBms.bFault OR i_stBms.bSystemLock));
// 2단계 BMS Minor(충전만 차단)와 통신 장애(15쪽: 정상운전 + 점검 요청)도 운전 단계는 멈추지만, 대기 단계에서는 기다림만
_bHardOk := _bDataOk AND NOT _bProtTrip AND NOT i_stUps.bBmsMinor;
// Rect Normal 0 = 정전·정류부 중고장(3단계) → 운전 단계 즉시 고장. BBC Normal은 BBC 기동 직후 3초 과도 구간에 0 → tModeTimeout 넘게 이어질 때만 고장
_bNormal := _bHardOk AND i_stUps.bRectNormal AND i_stUps.bBbcNormal;
_bActive := q_eStep <> E_UpsChargeStep.Idle AND q_eStep <> E_UpsChargeStep.WaitNormal
	AND q_eStep <> E_UpsChargeStep.Complete AND q_eStep <> E_UpsChargeStep.Fault;
// 스케줄 대기(최대 한 달)·휴지(30일)는 3~6단계만 고장. 그 밖의 이상은 고장으로 보지 않고 다음 단계로 넘어가지 않음
_bWaitStep := q_eStep = E_UpsChargeStep.WaitSchedule OR q_eStep = E_UpsChargeStep.Rest;
_tonAbnormal(IN:=_bActive AND NOT _bWaitStep AND _bHardOk AND i_stUps.bRectNormal AND NOT i_stUps.bBbcNormal,
	PT:=q_stActiveSet.tModeTimeout);
q_bConflict := q_eMode <> E_UpsChargeMode.Off AND i_eMode <> q_eMode AND i_eMode <> E_UpsChargeMode.Off;
IF i_bReset AND NOT i_bEnable AND (q_eStep = E_UpsChargeStep.Fault OR q_eStep = E_UpsChargeStep.Complete) THEN
	// 리셋은 현장 확인 후 수행. 장비를 정지시키는 명령이 아님.
	q_eStep := E_UpsChargeStep.Idle;
	q_eMode := E_UpsChargeMode.Off;
	q_nError := 0;
	q_bRecoveryRequired := FALSE;
	_bStarted := FALSE;
	_bSafeCancel := FALSE;
END_IF

IF _bActive THEN
	IF _bProtTrip OR (NOT _bWaitStep AND (NOT _bHardOk OR NOT i_stUps.bRectNormal OR _tonAbnormal.Q)) THEN
		_nNewFault := 2;
	ELSIF _fbRequest.q_bError THEN
		_nNewFault := 3;
	ELSIF NOT i_bEnable OR i_bCancel OR i_eMode = E_UpsChargeMode.Off THEN
		IF NOT _bCanceled THEN
			_bCanceled := TRUE;
			_bClearRequest := TRUE;
			IF NOT _bStarted THEN
				q_eStep := E_UpsChargeStep.Complete;
			ELSIF q_eMode = E_UpsChargeMode.Trickle THEN
				q_eStep := E_UpsChargeStep.BbcResume;
			ELSIF _bUpsDischargeRequested THEN
				q_eStep := E_UpsChargeStep.CancelUps;
			ELSE
				q_eStep := E_UpsChargeStep.CancelBms;
			END_IF
		END_IF
	END_IF
END_IF

_bEndReached := i_stUps.fBatteryVoltageV >= q_stActiveSet.fEndVoltageV;
_bRestartReached := i_stUps.fBatteryVoltageV <= q_stActiveSet.fStartVoltageV;
IF q_stActiveSet.nTrickleCriterion = 2 THEN
	_bEndReached := i_stBms.fSocPct >= q_stActiveSet.fEndSocPct;
	_bRestartReached := i_stBms.fSocPct <= q_stActiveSet.fStartSocPct;
END_IF
_tonExtra(IN:=q_eStep = E_UpsChargeStep.ExtraCharge, PT:=q_stActiveSet.tExtraCharge);
_tonRest(IN:=q_eStep = E_UpsChargeStep.Rest, PT:=q_stActiveSet.tRestart);
_tonInitial(IN:=q_eStep = E_UpsChargeStep.ExtraCharge AND q_eMode = E_UpsChargeMode.Periodic, PT:=q_stActiveSet.tInitialCharge);
_tonDischarge(IN:=q_eStep = E_UpsChargeStep.Running AND q_eMode = E_UpsChargeMode.Periodic, PT:=q_stActiveSet.tPeriodicDischarge);
_tonRun(IN:=q_eStep = E_UpsChargeStep.Running, PT:=q_stActiveSet.tRunTimeout);
_tonMode(IN:=q_eStep = E_UpsChargeStep.WaitRunning OR q_eStep = E_UpsChargeStep.WaitReady
	OR q_eStep = E_UpsChargeStep.WaitFloat, PT:=q_stActiveSet.tModeTimeout);
IF _nNewFault = 0 AND _tonMode.Q THEN _nNewFault:=4; END_IF
IF _nNewFault = 0 AND _tonRun.Q THEN _nNewFault:=5; END_IF
IF _nNewFault <> 0 THEN
	// UPS 방전을 요청하고 끝내지 못한 채 고장이면 방전 취소를 한 번 요청 (주기적 방전은 취소 전까지 계속됨)
	_bSafeCancel := _bUpsDischargeRequested AND (q_eStep = E_UpsChargeStep.StartDischarge
		OR q_eStep = E_UpsChargeStep.WaitRunning OR q_eStep = E_UpsChargeStep.Running OR q_eStep = E_UpsChargeStep.CancelUps);
	q_nError := _nNewFault;
	q_bRecoveryRequired := _bStarted OR _nNewFault = 5;
	_bClearRequest := TRUE; // 이전 요청의 확인·오류를 취소 요청에 다시 쓰지 않음
	q_eStep := E_UpsChargeStep.Fault;
END_IF

_bDue := FALSE;
IF i_stTime.bValid AND i_stTime.nMonth >= 1 AND i_stTime.nMonth <= 12
	AND i_stTime.nDay >= 1 AND i_stTime.nDay <= 31 THEN
	_nDate := UINT_TO_UDINT(i_stTime.nYear)*10000 + UINT_TO_UDINT(i_stTime.nMonth)*100 + UINT_TO_UDINT(i_stTime.nDay);
	_nWeek := (i_stTime.nDay-1)/7+1;
	_bDue := (q_stActiveSet.wMonthMask AND SHL(WORD#1,i_stTime.nMonth-1)) <> 0
		AND _nWeek = q_stActiveSet.nWeek AND i_stTime.nDayOfWeek = q_stActiveSet.nWeekDay
		AND i_stTime.nHour = q_stActiveSet.nHour AND _nDate > q_nLastScheduleDate;
END_IF

IF NOT _bClearRequest THEN
CASE q_eStep OF
	E_UpsChargeStep.Idle:
		IF i_bEnable AND NOT i_bCancel AND NOT i_bReset AND i_eMode <> E_UpsChargeMode.Off THEN
			q_eMode:=i_eMode; q_stActiveSet:=i_stSet; q_nError:=0;
			_bCanceled:=FALSE; _bStarted:=FALSE; _bUpsDischargeRequested:=FALSE;
			q_eStep:=E_UpsChargeStep.WaitNormal;
		END_IF
	E_UpsChargeStep.WaitNormal:
		IF NOT i_bEnable OR i_bCancel OR i_eMode = E_UpsChargeMode.Off THEN
			_bCanceled:=TRUE; q_eStep:=E_UpsChargeStep.Complete;
		ELSIF _bNormal THEN
			IF i_stUps.nBatMode <> 0 THEN
				q_bConflict:=TRUE;
			ELSIF q_stActiveSet.tRequestTimeout = T#0MS OR q_stActiveSet.tModeTimeout = T#0MS THEN
				q_nError:=1; q_eStep:=E_UpsChargeStep.Fault;
			ELSE
				CASE q_eMode OF
					E_UpsChargeMode.Trickle:
						IF (q_stActiveSet.nTrickleCriterion = 1 AND q_stActiveSet.fStartVoltageV > 0.0
							AND q_stActiveSet.fEndVoltageV > q_stActiveSet.fStartVoltageV)
							OR (q_stActiveSet.nTrickleCriterion = 2 AND q_stActiveSet.fStartSocPct >= 0.0
							AND q_stActiveSet.fEndSocPct > q_stActiveSet.fStartSocPct AND q_stActiveSet.fEndSocPct <= 100.0) THEN
							IF q_stActiveSet.tExtraCharge > T#0MS AND q_stActiveSet.tRestart > T#0MS THEN
								q_eStep:=E_UpsChargeStep.BbcStart;
							ELSE q_nError:=1; q_eStep:=E_UpsChargeStep.Fault; END_IF
						ELSE q_nError:=1; q_eStep:=E_UpsChargeStep.Fault; END_IF
					E_UpsChargeMode.Periodic:
						IF q_stActiveSet.fFloatVoltageV > 0.0 AND q_stActiveSet.fPeriodicCurrentA > 0.0
							AND q_stActiveSet.tInitialCharge > T#0MS AND q_stActiveSet.tPeriodicDischarge > T#0MS AND q_stActiveSet.tRunTimeout > q_stActiveSet.tPeriodicDischarge
							AND q_stActiveSet.wMonthMask <> 0 AND q_stActiveSet.wMonthMask <= 16#0FFF
							AND q_stActiveSet.nWeek >= 1 AND q_stActiveSet.nWeek <= 4
							AND q_stActiveSet.nWeekDay <= 6 AND q_stActiveSet.nHour <= 23 THEN
							q_eStep:=E_UpsChargeStep.WaitSchedule;
						ELSE q_nError:=1; q_eStep:=E_UpsChargeStep.Fault; END_IF
					E_UpsChargeMode.Pulse:
						IF q_stActiveSet.fPulseChargeA > 0.0 AND q_stActiveSet.fPulseDischargeA > 0.0
							AND q_stActiveSet.tPulseCharge > T#0MS AND q_stActiveSet.tPulseDischarge > T#0MS
							AND q_stActiveSet.nPulseCycles > 0 AND q_stActiveSet.tRunTimeout > T#0MS
							AND (UDINT_TO_LREAL(TIME_TO_UDINT(q_stActiveSet.tPulseCharge))
							+ UDINT_TO_LREAL(TIME_TO_UDINT(q_stActiveSet.tPulseDischarge)))
							*UINT_TO_LREAL(q_stActiveSet.nPulseCycles) < UDINT_TO_LREAL(TIME_TO_UDINT(q_stActiveSet.tRunTimeout)) THEN
							q_eStep:=E_UpsChargeStep.PrepareBms;
						ELSE q_nError:=1; q_eStep:=E_UpsChargeStep.Fault; END_IF
					ELSE q_nError:=1; q_eStep:=E_UpsChargeStep.Fault;
				END_CASE
			END_IF
		END_IF
	E_UpsChargeStep.WaitSchedule:
		IF _bDue AND i_stUps.nBatMode = 0 AND _bNormal THEN
			q_nLastScheduleDate:=_nDate;
			IF i_stUps.fBatteryVoltageV <= q_stActiveSet.fFloatVoltageV THEN q_eStep:=E_UpsChargeStep.ExtraCharge;
			ELSE q_eStep:=E_UpsChargeStep.PrepareBms; END_IF
		END_IF
	E_UpsChargeStep.BbcStart:
		IF _fbRequest.q_bDone THEN q_eStep:=E_UpsChargeStep.WaitEnd;
		ELSE _eAction:=E_UpsChargeAction.BbcOn; _bStarted:=TRUE; END_IF
	E_UpsChargeStep.WaitEnd:
		IF _bEndReached THEN q_eStep:=E_UpsChargeStep.ExtraCharge; END_IF
	E_UpsChargeStep.ExtraCharge:
		IF q_eMode = E_UpsChargeMode.Trickle AND _tonExtra.Q THEN q_eStep:=E_UpsChargeStep.BbcReady;
		ELSIF q_eMode = E_UpsChargeMode.Periodic AND _tonInitial.Q THEN q_eStep:=E_UpsChargeStep.PrepareBms; END_IF
	E_UpsChargeStep.BbcReady:
		IF _fbRequest.q_bDone THEN _nModeSample:=i_stUps.nSampleSeq; q_eStep:=E_UpsChargeStep.WaitReady;
		ELSE _eAction:=E_UpsChargeAction.BbcReady; END_IF
	E_UpsChargeStep.WaitReady:
		IF i_stUps.nSampleSeq <> _nModeSample AND i_stUps.nBatMode = 2 THEN q_eStep:=E_UpsChargeStep.Rest; END_IF
	E_UpsChargeStep.Rest:
		IF (_bRestartReached OR _tonRest.Q) AND _bHardOk AND i_stUps.bRectNormal THEN q_eStep:=E_UpsChargeStep.BbcStart; END_IF // 대기모드에서는 BBC Normal을 보지 않음
	E_UpsChargeStep.PrepareBms:
		IF i_stUps.nBatMode <> 0 THEN q_bConflict:=TRUE;
		ELSIF _fbRequest.q_bDone THEN q_eStep:=E_UpsChargeStep.StartDischarge;
		ELSE
			_bStarted:=TRUE;
			IF q_eMode = E_UpsChargeMode.Periodic THEN _eAction:=E_UpsChargeAction.BmsPreparePeriodic;
			ELSE _eAction:=E_UpsChargeAction.BmsPreparePulse; END_IF
		END_IF
	E_UpsChargeStep.StartDischarge:
		IF NOT _bUpsDischargeRequested AND i_stUps.nBatMode <> 0 THEN q_bConflict:=TRUE;
		ELSIF _fbRequest.q_bDone THEN _nModeSample:=i_stUps.nSampleSeq; q_eStep:=E_UpsChargeStep.WaitRunning;
		ELSE
			_bUpsDischargeRequested:=TRUE;
			IF q_eMode = E_UpsChargeMode.Periodic THEN _eAction:=E_UpsChargeAction.PeriodicStart;
			ELSE _eAction:=E_UpsChargeAction.PulseStart; END_IF
		END_IF
	E_UpsChargeStep.WaitRunning:
		IF i_stUps.nSampleSeq <> _nModeSample AND ((q_eMode = E_UpsChargeMode.Periodic AND i_stUps.nBatMode = 3)
			OR (q_eMode = E_UpsChargeMode.Pulse AND i_stUps.nBatMode = 4)) THEN
			q_fStartVoltageV:=i_stUps.fBatteryVoltageV;
			_nModeSample:=i_stUps.nSampleSeq; q_eStep:=E_UpsChargeStep.Running;
		END_IF
	E_UpsChargeStep.Running:
		IF (q_eMode = E_UpsChargeMode.Periodic AND i_stUps.nBatMode = 3) OR (q_eMode = E_UpsChargeMode.Pulse AND i_stUps.nBatMode = 4) THEN
			q_fEndVoltageV:=i_stUps.fBatteryVoltageV; // 방전 중 마지막 전압 = 종료 전압 (부동충전 복귀 뒤에는 전압이 다시 오름)
		END_IF
		IF i_stUps.nSampleSeq <> _nModeSample AND i_stUps.nBatMode = 0 THEN q_eStep:=E_UpsChargeStep.CancelBms;
		ELSIF q_eMode = E_UpsChargeMode.Periodic AND _tonDischarge.Q THEN q_eStep:=E_UpsChargeStep.CancelUps; END_IF
	E_UpsChargeStep.CancelUps:
		IF _fbRequest.q_bDone THEN q_eStep:=E_UpsChargeStep.CancelBms;
		ELSE _eAction:=E_UpsChargeAction.DischargeCancel; END_IF
	E_UpsChargeStep.CancelBms:
		IF _fbRequest.q_bDone THEN q_eStep:=E_UpsChargeStep.FloatRequest;
		ELSE _eAction:=E_UpsChargeAction.BmsDischargeCancel; END_IF
	E_UpsChargeStep.BbcResume:
		IF _fbRequest.q_bDone THEN q_eStep:=E_UpsChargeStep.FloatRequest;
		ELSE _eAction:=E_UpsChargeAction.BbcOn; END_IF
	E_UpsChargeStep.FloatRequest:
		IF _fbRequest.q_bDone THEN _nModeSample:=i_stUps.nSampleSeq; q_eStep:=E_UpsChargeStep.WaitFloat;
		ELSE _eAction:=E_UpsChargeAction.FloatCharge; END_IF
	E_UpsChargeStep.WaitFloat:
		IF i_stUps.nSampleSeq <> _nModeSample AND i_stUps.nBatMode = 0 THEN
			IF q_eMode = E_UpsChargeMode.Trickle THEN q_fEndVoltageV:=i_stUps.fBatteryVoltageV; END_IF
			q_stLastTime:=i_stTime; _bStarted:=FALSE; _bUpsDischargeRequested:=FALSE;
			IF _bCanceled THEN q_eStep:=E_UpsChargeStep.Complete;
			ELSIF q_eMode = E_UpsChargeMode.Periodic THEN
				IF NOT q_bReferenceValid THEN
					q_fReferenceStartVoltageV:=q_fStartVoltageV;
					q_fReferenceEndVoltageV:=q_fEndVoltageV;
					q_stReferenceTime:=i_stTime; q_bReferenceValid:=TRUE;
				END_IF
				q_bDone:=TRUE; q_eStep:=E_UpsChargeStep.WaitSchedule;
			ELSE q_bDone:=TRUE; q_eStep:=E_UpsChargeStep.Complete; END_IF
		END_IF
	E_UpsChargeStep.Complete:
		q_bCanceled:=_bCanceled;
		IF NOT i_bEnable THEN q_eStep:=E_UpsChargeStep.Idle; q_eMode:=E_UpsChargeMode.Off; END_IF
	E_UpsChargeStep.Fault:
		// 장비 보호·비상정지는 별도 담당. 자동 재시작하지 않음. 방전 중이었으면 UPS 데이터가 유효할 때 취소를 한 번 요청
		IF _bSafeCancel THEN
			IF _fbRequest.q_bDone OR _fbRequest.q_bError THEN _bSafeCancel:=FALSE;
			ELSIF i_stUps.bValid THEN _eAction:=E_UpsChargeAction.DischargeCancel; END_IF
		END_IF
END_CASE
END_IF
_fbRequest(i_eAction:=_eAction, i_fValue:=0.0, i_tTimeout:=q_stActiveSet.tRequestTimeout, i_stFeedback:=i_stFeedback);
q_stRequest:=_fbRequest.q_stRequest;

END_FUNCTION_BLOCK

// ---- 20_Module/Ups/FB_UpsTemperatureCharge.TcPOU
FUNCTION_BLOCK FB_UpsTemperatureCharge // 온도보상 전압 계산 및 적용 요청
VAR_INPUT
	i_bEnable : BOOL;
	i_bSuspend : BOOL;
	i_bReset : BOOL;
	i_stUps : ST_UpsState;
	i_stSet : ST_UpsChargeSet;
	i_stTime : ST_LocalTime;
	i_stFeedback : ST_UpsChargeFeedback;
END_VAR
VAR_OUTPUT
	q_stRequest : ST_UpsChargeRequest;
	q_fTargetVoltageV : REAL;
	q_fAppliedVoltageV : REAL;
	q_bSuspended : BOOL;
	q_bApplied : BOOL;
	q_nError : UINT; // 1: 설정/온도, 2: 통신/보호, 3: 적용 확인
	q_stLastTime : ST_LocalTime;
END_VAR
VAR
	_fbRequest : FB_UpsChargeRequest;
	_eAction : E_UpsChargeAction;
	_tonUpdate : TON;
	_bUpdateDone : BOOL;
	_bRestore : BOOL;
	_bWasSuspended : BOOL;
	_fPendingV : REAL;
	_bPending : BOOL;
END_VAR

_eAction:=E_UpsChargeAction.NoRequest;
q_bSuspended:=i_bSuspend OR i_stUps.nBatMode = 3 OR i_stUps.nBatMode = 4;
_tonUpdate(IN:=q_bApplied AND NOT _bUpdateDone, PT:=i_stSet.tTempUpdate);
_bUpdateDone:=FALSE;
IF i_bReset THEN q_nError:=0; END_IF
IF q_nError = 2 THEN q_nError:=0; END_IF // 통신·보호 이상은 래치하지 않음: 매 스캔 다시 판정, 풀리면 이어서 (Disable이면 부동충전 전압 복귀)
IF _fbRequest.q_bError THEN q_nError:=3; END_IF

IF q_nError = 0 AND (i_bEnable OR q_bApplied OR _bPending) THEN
	IF NOT i_stUps.bValid OR NOT i_stUps.bRectNormal OR NOT i_stUps.bBbcNormal
		OR i_stUps.bEmergencyStop OR i_stUps.bBmsMinor OR i_stUps.bBmsMajor
		OR (i_stUps.wStatus2 AND 16#7000) <> 0 OR (i_stUps.wBbcAlarm AND 16#0FA8) <> 0 THEN // RCD 1·2단계·화재, BBC 정지 알람 (동작시퀀스 7쪽)
		q_nError:=2; _bPending:=FALSE;
	ELSIF NOT (i_stSet.fBaseCellVoltageV > 0.0 AND i_stSet.nSeriesCells > 0
		AND i_stSet.fMinChargeVoltageV > 0.0
		AND i_stSet.fMaxChargeVoltageV >= i_stSet.fMinChargeVoltageV
		AND i_stSet.fMaxChargeVoltageV <= 6553.5
		AND i_stSet.fFloatVoltageV >= i_stSet.fMinChargeVoltageV
		AND i_stSet.fFloatVoltageV <= i_stSet.fMaxChargeVoltageV
		AND i_stSet.fMinTemperatureC < i_stSet.fMaxTemperatureC
		AND i_stSet.tRequestTimeout > T#0MS AND i_stSet.tTempUpdate > T#0MS) THEN
		q_nError:=1;
	ELSIF NOT q_bSuspended THEN
		IF NOT _bPending THEN
			_bRestore:=NOT i_bEnable;
			IF _bRestore THEN q_fTargetVoltageV:=i_stSet.fFloatVoltageV;
			ELSE
				IF i_stUps.fBatteryRoomTemperatureC < i_stSet.fMinTemperatureC
					OR i_stUps.fBatteryRoomTemperatureC > i_stSet.fMaxTemperatureC THEN q_nError:=1;
				ELSE q_fTargetVoltageV:=(i_stSet.fBaseCellVoltageV + i_stSet.fSlopeMvPerC*0.001
					*(i_stUps.fBatteryRoomTemperatureC-25.0))*UINT_TO_REAL(i_stSet.nSeriesCells); END_IF
			END_IF
			IF NOT (q_fTargetVoltageV >= i_stSet.fMinChargeVoltageV AND q_fTargetVoltageV <= i_stSet.fMaxChargeVoltageV) THEN q_nError:=1; END_IF
			// 주기 갱신은 전압이 레지스터 해상도(0.1 V) 이상 바뀔 때만 씀. 아니면 쓰지 않고 주기만 다시 시작
			IF q_nError = 0 AND (NOT q_bApplied OR _bRestore OR _bWasSuspended
				OR (_tonUpdate.Q AND ABS(q_fTargetVoltageV - q_fAppliedVoltageV) >= 0.1)) THEN
				_fPendingV:=q_fTargetVoltageV; _bPending:=TRUE;
			ELSIF _tonUpdate.Q THEN
				_bUpdateDone:=TRUE;
			END_IF
		END_IF
		IF _bPending AND q_nError = 0 THEN
			IF _fbRequest.q_bDone THEN
				q_fAppliedVoltageV:=_fPendingV; q_stLastTime:=i_stTime;
				q_bApplied:=NOT _bRestore; _bPending:=FALSE; _bUpdateDone:=TRUE;
			ELSE _eAction:=E_UpsChargeAction.ChargeVoltage; END_IF
		END_IF
	END_IF
END_IF
IF q_bSuspended THEN _bPending:=FALSE; END_IF
_bWasSuspended:=q_bSuspended;
_fbRequest(i_eAction:=_eAction, i_fValue:=_fPendingV, i_tTimeout:=i_stSet.tRequestTimeout, i_stFeedback:=i_stFeedback);
q_stRequest:=_fbRequest.q_stRequest;

END_FUNCTION_BLOCK

